(* IEC 61131-3 sources: plc-st-coding-agent/progress/evidence/f14_v10_full_20261113/jobs/codex_minimax-m27 (part 5) *)

(* ---- public-medium-04.candidate_04.st ---- *)
(* CONTRACT_RULES [] *)
FUNCTION_BLOCK FB_TemperatureControl
VAR_INPUT
    TemperatureSensorInput : REAL;
    SetTemperature         : REAL;
END_VAR
VAR_OUTPUT
    CurrentTemperature : REAL;
    SetTempDisplay      : REAL;
    HeaterStatus        : BOOL;
    OverheatProtection  : BOOL;
    HeaterOutput        : BOOL;
END_VAR
VAR
    tonCooldown         : TON;
    local_OverheatActive : BOOL := FALSE;
    local_SensorFault    : BOOL := FALSE;
    local_RuntimeAccum   : LTIME := LTIME#0s;
END_VAR

(* ENGINEERING_CONTRACT
  PUB003: Overheat protection triggers when heater runs continuously > 5s.
    - Activation: local_RuntimeAccum exceeds 5s on same scan it is detected.
    - Retention: OverheatActive stays TRUE until cooldown completes.
    - Reset/Deactivation: 3s cooldown via tonCooldown; heating condition
      must reassert AND cooldown must complete before heater can restart.
    - Same-scan priority: heater outputs set to FALSE when overheat activates;
      local_RuntimeAccum resets only when heating condition drops (not on
      overheat trigger), preserving correct accumulated-time logic.
    - Units/Boundaries: LTIME nanoseconds; strict > 5000ms threshold.
  PUB004: Heater turns on when temperature < setpoint (strict <).
  PUB007: Status outputs reflect current state every scan.
  PUB006: Sensor fault (input < 0 or > 100) turns heater off immediately.
*)

CurrentTemperature := TemperatureSensorInput;
SetTempDisplay     := SetTemperature;

local_SensorFault := (TemperatureSensorInput < 0.0) OR (TemperatureSensorInput > 100.0);

IF local_SensorFault OR local_OverheatActive THEN
    HeaterOutput := FALSE;
ELSE
    IF TemperatureSensorInput < SetTemperature THEN
        HeaterOutput := TRUE;
    ELSE
        HeaterOutput := FALSE;
    END_IF;
END_IF;

IF HeaterOutput THEN
    local_RuntimeAccum := local_RuntimeAccum + TO_LTIME(1);
END_IF;

IF NOT HeaterOutput THEN
    local_RuntimeAccum := LTIME#0s;
END_IF;

IF local_RuntimeAccum > T#5s THEN
    local_OverheatActive := TRUE;
    local_RuntimeAccum   := LTIME#0s;
END_IF;

IF local_OverheatActive THEN
    tonCooldown(IN := TRUE, PT := T#3s);
    IF tonCooldown.Q THEN
        local_OverheatActive := FALSE;
    END_IF;
ELSE
    tonCooldown(IN := FALSE, PT := T#3s);
END_IF;

HeaterStatus       := HeaterOutput;
OverheatProtection := local_OverheatActive;
END_FUNCTION_BLOCK

(* ---- public-medium-04.raw_candidate_01.st ---- *)
(*
ENGINEERING_CONTRACT:
PUB001: Read TemperatureSensorInput (REAL), display in CurrentTemperature
PUB002: HeaterOutput := TRUE when TemperatureSensorInput < SetTemperature
PUB003: Overheat triggers after >5s continuous HeaterOutput (strict > boundary)
PUB004: Overheat auto-sets HeaterOutput:=FALSE, 3s cooldown before OverheatProtection can clear
PUB005: Sensor fault (<0 OR >100) sets HeaterOutput:=FALSE regardless of temperature
PUB006: Status outputs (CurrentTemperature, SetTempDisplay, HeaterStatus, OverheatProtection) update every scan

Activation: All outputs update every scan (no edge-only behavior)
Retention: OverheatActive retains state across scans until cooldown completes
Reset/Deactivation: OverheatActive resets only after OverheatCooldownTimer.Q (3s elapsed)
Same-scan priority: HeaterOutput finalized BEFORE runtime timer enable is evaluated
Units: TIME/LTIME for timers (TON), REAL for temperatures, BOOL for control/status
*)
FUNCTION_BLOCK FB_TemperatureControl
VAR_INPUT
    TemperatureSensorInput : REAL;
    SetTemperature : REAL;
END_VAR

VAR_OUTPUT
    CurrentTemperature : REAL;
    SetTempDisplay : REAL;
    HeaterStatus : BOOL;
    OverheatProtection : BOOL;
    HeaterOutput : BOOL;
END_VAR

VAR
    HeaterRuntimeTimer : TON;
    OverheatCooldownTimer : TON;
    OverheatActive : BOOL := FALSE;
    SensorFault : BOOL := FALSE;
END_VAR

// Update display outputs
CurrentTemperature := TemperatureSensorInput;
SetTempDisplay := SetTemperature;

// Sensor fault detection: invalid range turns off heater
SensorFault := (TemperatureSensorInput < 0.0) OR (TemperatureSensorInput > 100.0);

// Temperature control logic
IF NOT SensorFault AND NOT OverheatActive THEN
    // Normal operation: heater ON when below setpoint
    IF TemperatureSensorInput < SetTemperature THEN
        HeaterOutput := TRUE;
    ELSE
        HeaterOutput := FALSE;
    END_IF;
ELSE
    // Sensor fault or overheat protection active - heater OFF
    HeaterOutput := FALSE;
END_IF;

// Update heater status display
HeaterStatus := HeaterOutput;

// Runtime timer: tracks continuous heater ON time (resets when heater OFF)
HeaterRuntimeTimer(IN := HeaterOutput, PT := T#5s);

// Overheat detection: >5s continuous heater operation
IF HeaterRuntimeTimer.Q AND NOT OverheatActive THEN
    OverheatActive := TRUE;
    OverheatCooldownTimer(IN := TRUE, PT := T#3s);
END_IF;

// Overheat cooldown: 3s wait before protection can be lifted
IF OverheatActive THEN
    OverheatCooldownTimer(IN := TRUE, PT := T#3s);
    IF OverheatCooldownTimer.Q THEN
        OverheatActive := FALSE;
    END_IF;
END_IF;

// Update overheat protection status
OverheatProtection := OverheatActive;
END_FUNCTION_BLOCK

(* ---- public-medium-04.raw_candidate_02.st ---- *)
(*
ENGINEERING_CONTRACT:
PUB001: TemperatureSensorInput (REAL) -> CurrentTemperature (REAL) every scan
PUB002: HeaterOutput := TRUE when TemperatureSensorInput < SetTemperature (no sensor fault)
PUB003: Overheat triggers when runtime > 5s (strict >), first satisfying tick = 5001ms
PUB004: Overheat sets HeaterOutput:=FALSE, 3s cooldown before OverheatProtection clears
PUB005: Sensor fault (<0 OR >100) sets HeaterOutput:=FALSE regardless of temperature
PUB006: All status outputs (CurrentTemperature, SetTempDisplay, HeaterStatus, OverheatProtection) update every scan
*)
FUNCTION_BLOCK FB_TemperatureControl
VAR_INPUT
    TemperatureSensorInput : REAL;
    SetTemperature         : REAL;
END_VAR

VAR_OUTPUT
    CurrentTemperature : REAL;
    SetTempDisplay      : REAL;
    HeaterStatus        : BOOL;
    OverheatProtection  : BOOL;
    HeaterOutput        : BOOL;
END_VAR

VAR
    HeaterRuntimeTimer   : TON;
    OverheatCooldownTimer: TON;
    OverheatActive       : BOOL := FALSE;
    SensorFault          : BOOL := FALSE;
    Runtimems            : LINT := 0;
END_VAR

SensorFault := (TemperatureSensorInput < 0.0) OR (TemperatureSensorInput > 100.0);

IF NOT SensorFault AND NOT OverheatActive THEN
    IF TemperatureSensorInput < SetTemperature THEN
        HeaterOutput := TRUE;
    ELSE
        HeaterOutput := FALSE;
    END_IF;
ELSE
    HeaterOutput := FALSE;
END_IF;

HeaterRuntimeTimer(IN := FALSE, PT := T#5s);

IF OverheatActive THEN
    IF Runtimems > 5000 THEN
        OverheatActive := TRUE;
    END_IF;
ELSIF HeaterOutput THEN
    Runtimems := Runtimems + TO_LINT(HeaterRuntimeTimer.ET) + 1;
    HeaterRuntimeTimer(IN := TRUE, PT := T#5s);
    IF Runtimems > 5000 THEN
        OverheatActive := TRUE;
        HeaterOutput := FALSE;
    END_IF;
ELSE
    Runtimems := 0;
END_IF;

IF OverheatActive THEN
    OverheatCooldownTimer(IN := TRUE, PT := T#3s);
    IF OverheatCooldownTimer.Q THEN
        OverheatActive := FALSE;
        Runtimems := 0;
    END_IF;
END_IF;

CurrentTemperature := TemperatureSensorInput;
SetTempDisplay := SetTemperature;
HeaterStatus := HeaterOutput;
OverheatProtection := OverheatActive;
END_FUNCTION_BLOCK

(* ---- public-medium-04.raw_candidate_03.st ---- *)
(* CONTRACT_RULES [] *)
FUNCTION_BLOCK FB_TemperatureControl
VAR_INPUT
    TemperatureSensorInput : REAL;
    SetTemperature : REAL;
END_VAR
VAR_OUTPUT
    CurrentTemperature : REAL;
    SetTempDisplay : REAL;
    HeaterStatus : BOOL;
    OverheatProtection : BOOL;
    HeaterOutput : BOOL;
END_VAR
VAR
    HeaterRuntimeTimer : TON;
    OverheatCooldownTimer : TON;
    OverheatActive : BOOL := FALSE;
    SensorFault : BOOL := FALSE;
END_VAR

CurrentTemperature := TemperatureSensorInput;
SetTempDisplay := SetTemperature;
SensorFault := (TemperatureSensorInput < 0.0) OR (TemperatureSensorInput > 100.0);

HeaterRuntimeTimer(IN := (TemperatureSensorInput < SetTemperature) AND NOT SensorFault AND NOT OverheatActive, PT := T#5s);

IF HeaterRuntimeTimer.Q AND NOT OverheatActive THEN
    OverheatActive := TRUE;
    OverheatCooldownTimer(IN := TRUE, PT := T#3s);
END_IF;

IF OverheatActive THEN
    OverheatCooldownTimer(IN := TRUE, PT := T#3s);
    IF OverheatCooldownTimer.Q THEN
        OverheatActive := FALSE;
    END_IF;
END_IF;

IF NOT SensorFault AND NOT OverheatActive THEN
    IF TemperatureSensorInput < SetTemperature THEN
        HeaterOutput := TRUE;
    ELSE
        HeaterOutput := FALSE;
    END_IF;
ELSE
    HeaterOutput := FALSE;
END_IF;

HeaterStatus := HeaterOutput;
OverheatProtection := OverheatActive;
END_FUNCTION_BLOCK

(* ---- public-medium-04.raw_candidate_04.st ---- *)
(* CONTRACT_RULES [] *)
FUNCTION_BLOCK FB_TemperatureControl
VAR_INPUT
    TemperatureSensorInput : REAL;
    SetTemperature         : REAL;
END_VAR
VAR_OUTPUT
    CurrentTemperature : REAL;
    SetTempDisplay      : REAL;
    HeaterStatus        : BOOL;
    OverheatProtection  : BOOL;
    HeaterOutput        : BOOL;
END_VAR
VAR
    tonCooldown         : TON;
    local_OverheatActive : BOOL := FALSE;
    local_SensorFault    : BOOL := FALSE;
    local_RuntimeAccum   : LTIME := LTIME#0s;
END_VAR

(* ENGINEERING_CONTRACT
  PUB003: Overheat protection triggers when heater runs continuously > 5s.
    - Activation: local_RuntimeAccum exceeds 5s on same scan it is detected.
    - Retention: OverheatActive stays TRUE until cooldown completes.
    - Reset/Deactivation: 3s cooldown via tonCooldown; heating condition
      must reassert AND cooldown must complete before heater can restart.
    - Same-scan priority: heater outputs set to FALSE when overheat activates;
      local_RuntimeAccum resets only when heating condition drops (not on
      overheat trigger), preserving correct accumulated-time logic.
    - Units/Boundaries: LTIME nanoseconds; strict > 5000ms threshold.
  PUB004: Heater turns on when temperature < setpoint (strict <).
  PUB007: Status outputs reflect current state every scan.
  PUB006: Sensor fault (input < 0 or > 100) turns heater off immediately.
*)

CurrentTemperature := TemperatureSensorInput;
SetTempDisplay     := SetTemperature;

local_SensorFault := (TemperatureSensorInput < 0.0) OR (TemperatureSensorInput > 100.0);

IF local_SensorFault OR local_OverheatActive THEN
    HeaterOutput := FALSE;
ELSE
    IF TemperatureSensorInput < SetTemperature THEN
        HeaterOutput := TRUE;
    ELSE
        HeaterOutput := FALSE;
    END_IF;
END_IF;

IF HeaterOutput THEN
    local_RuntimeAccum := local_RuntimeAccum + TO_LTIME(1);
END_IF;

IF NOT HeaterOutput THEN
    local_RuntimeAccum := LTIME#0s;
END_IF;

IF local_RuntimeAccum > T#5s THEN
    local_OverheatActive := TRUE;
    local_RuntimeAccum   := LTIME#0s;
END_IF;

IF local_OverheatActive THEN
    tonCooldown(IN := TRUE, PT := T#3s);
    IF tonCooldown.Q THEN
        local_OverheatActive := FALSE;
    END_IF;
ELSE
    tonCooldown(IN := FALSE, PT := T#3s);
END_IF;

HeaterStatus       := HeaterOutput;
OverheatProtection := local_OverheatActive;
END_FUNCTION_BLOCK

(* ---- public-medium-05.candidate_01.st ---- *)
(* ENGINEERING_CONTRACT *)
(*
  | Output/State Group       | Activation                                  | Retention                    | Reset/Deactivation            | Same-Scan Priority | Units/Boundaries |
  |--------------------------|---------------------------------------------|------------------------------|-------------------------------|--------------------|------------------|
  | MotorForward (Auto)      | State<>IDLE AND Mode=1                      | Hold until State=IDLE        | State=IDLE OR Mode=0          | Same-scan          | PUB001,PUB007    |
  | MotorReverse (Manual)    | ForwardButton=1 AND Mode=0 AND ReverseButton=0 | Hold until condition false | ForwardButton=0 OR Mode=1   | Same-scan          | PUB006,PUB002    |
  | CompletionLight          | State=DONE AND SensorC=1 AND Mode=1         | Hold while SensorC=1         | SensorC=0 OR Mode=0           | Same-scan          | PUB004,PUB008    |
  | State: IDLE→A            | SensorA=1 AND Mode=1 AND State=IDLE         | Until next transition        | SensorC=0 (product removed)   | Same-scan          | PUB003           |
  | State: A→B               | ButtonA=1 AND State=A                       | Until next transition        | SensorC=0                      | Same-scan          | PUB003           |
  | State: B→C               | SensorB=1 AND State=B                       | Until next transition        | SensorC=0                      | Same-scan          | PUB003           |
  | State: C→DONE            | ButtonC=1 AND State=C                       | Until SensorC=0              | SensorC=0                      | Same-scan          | PUB003           |
*)
(* CONTRACT_RULES [] *)
FUNCTION_BLOCK ProductionLineControl
VAR_INPUT
    Mode : BOOL;
    ForwardButton : BOOL;
    ReverseButton : BOOL;
    SensorA : BOOL;
    SensorB : BOOL;
    SensorC : BOOL;
    ButtonA : BOOL;
    ButtonB : BOOL;
    ButtonC : BOOL;
END_VAR
VAR_OUTPUT
    MotorForward : BOOL;
    MotorReverse : BOOL;
    CompletionLight : BOOL;
END_VAR
VAR
    State : INT;
    IDLE : INT := 0;
    StateA : INT := 1;
    StateB : INT := 2;
    StateC : INT := 3;
    StateD : INT := 4;
END_VAR
    IF Mode = FALSE THEN
        State := IDLE;
    ELSIF Mode = TRUE THEN
        IF State = IDLE AND SensorA THEN
            State := StateA;
        ELSIF State = StateA AND ButtonA THEN
            State := StateB;
        ELSIF State = StateB AND SensorB THEN
            State := StateC;
        ELSIF State = StateC AND ButtonC THEN
            State := StateD;
        END_IF;
    END_IF;
    MotorForward := ((State <> IDLE) AND Mode) OR (ForwardButton AND (NOT Mode) AND (NOT ReverseButton));
    MotorReverse := ReverseButton AND (NOT Mode) AND (NOT ForwardButton);
    CompletionLight := (State = StateD) AND SensorC AND Mode;
END_FUNCTION_BLOCK

(* ---- public-medium-05.candidate_02.st ---- *)
(* ENGINEERING_CONTRACT *)
(*
  | Output/State Group       | Activation                                  | Retention                    | Reset/Deactivation            | Same-Scan Priority | Units/Boundaries |
  |--------------------------|---------------------------------------------|------------------------------|-------------------------------|--------------------|------------------|
  | MotorForward (Auto)      | State=B OR State=D_transit                  | Hold via tmp_MotorRunning    | State=C/DONE OR Mode=0         | Same-scan          | PUB006           |
  | MotorReverse (Manual)    | ReverseButton AND Mode=0 AND !ForwardButton | Hold until condition false   | !ReverseButton OR Mode=1       | Same-scan          | PUB004,PUB002    |
  | CompletionLight          | State=DONE AND SensorC AND Mode             | Hold while SensorC           | SensorC=0 OR Mode=0            | Same-scan          | PUB008           |
  | State transitions        | Per clause PUB003                           | Until next trigger           | Mode=0 → IDLE                  | Same-scan          | PUB003           |
*)
(* CONTRACT_RULES [] *)
FUNCTION_BLOCK ProductionLineControl
VAR_INPUT
    Mode : BOOL;
    ForwardButton : BOOL;
    ReverseButton : BOOL;
    SensorA : BOOL;
    SensorB : BOOL;
    SensorC : BOOL;
    ButtonA : BOOL;
    ButtonB : BOOL;
    ButtonC : BOOL;
END_VAR
VAR_OUTPUT
    MotorForward : BOOL;
    MotorReverse : BOOL;
    CompletionLight : BOOL;
END_VAR
VAR
    State : INT;
    IDLE : INT := 0;
    StateA : INT := 1;
    StateB : INT := 2;
    StateC : INT := 3;
    StateD_transit : INT := 4;
    DONE : INT := 5;
    tmp_MotorRunning : BOOL;
END_VAR
    tmp_MotorRunning := (State = StateB) OR (State = StateD_transit);
    MotorForward := tmp_MotorRunning AND Mode;
    MotorReverse := ReverseButton AND (NOT Mode) AND (NOT ForwardButton);
    CompletionLight := (State = DONE) AND SensorC AND Mode;
    IF Mode = FALSE THEN
        State := IDLE;
    ELSIF Mode = TRUE THEN
        IF State = IDLE AND SensorA THEN
            State := StateA;
        ELSIF State = StateA AND ButtonA THEN
            State := StateB;
            tmp_MotorRunning := TRUE;
        ELSIF State = StateB AND SensorB THEN
            State := StateC;
        ELSIF State = StateC AND ButtonC THEN
            State := StateD_transit;
            tmp_MotorRunning := TRUE;
        ELSIF State = StateD_transit AND SensorC THEN
            State := DONE;
        ELSIF State = DONE AND NOT SensorC THEN
            State := IDLE;
        END_IF;
    END_IF;
END_FUNCTION_BLOCK

(* ---- public-medium-05.candidate_03.st ---- *)
(* ENGINEERING_CONTRACT *)
(*
  | Output/State Group       | Activation                                  | Retention                    | Reset/Deactivation            | Same-Scan Priority | Units/Boundaries |
  |--------------------------|---------------------------------------------|------------------------------|-------------------------------|--------------------|------------------|
  | MotorForward (Auto)      | State=StateA OR State=StateB AND Mode=1      | Hold until State=C or IDLE   | State=C/D OR Mode=0          | Same-scan          | PUB001,PUB007    |
  | MotorReverse (Manual)    | ForwardButton=1 AND Mode=0 AND ReverseButton=0 | Hold until condition false | ForwardButton=0 OR Mode=1   | Same-scan          | PUB006,PUB002    |
  | CompletionLight          | State=StateD AND SensorC=1 AND Mode=1        | Hold while SensorC=1         | SensorC=0 OR Mode=0           | Same-scan          | PUB004,PUB008    |
  | State: IDLE→A            | SensorA=1 AND Mode=1 AND State=IDLE          | Until next transition        | SensorC=0 (product removed)   | Same-scan          | PUB003           |
  | State: A→B               | ButtonA=1 AND State=StateA                   | Until next transition        | SensorC=0                     | Same-scan          | PUB003           |
  | State: B→C               | SensorB=1 AND State=StateB                   | Until next transition        | SensorC=0                     | Same-scan          | PUB003           |
  | State: C→DONE            | ButtonC=1 AND State=StateC                   | Until SensorC=0              | SensorC=0                     | Same-scan          | PUB003           |
*)
(* CONTRACT_RULES [] *)
FUNCTION_BLOCK ProductionLineControl
VAR_INPUT
    Mode : BOOL;
    ForwardButton : BOOL;
    ReverseButton : BOOL;
    SensorA : BOOL;
    SensorB : BOOL;
    SensorC : BOOL;
    ButtonA : BOOL;
    ButtonB : BOOL;
    ButtonC : BOOL;
END_VAR
VAR_OUTPUT
    MotorForward : BOOL;
    MotorReverse : BOOL;
    CompletionLight : BOOL;
END_VAR
VAR
    State : INT;
    IDLE : INT := 0;
    StateA : INT := 1;
    StateB : INT := 2;
    StateC : INT := 3;
    StateD : INT := 4;
END_VAR
    IF Mode = FALSE THEN
        State := IDLE;
    ELSIF Mode = TRUE THEN
        IF State = IDLE AND SensorA THEN
            State := StateA;
        ELSIF State = StateA AND ButtonA THEN
            State := StateB;
        ELSIF State = StateB AND SensorB THEN
            State := StateC;
        ELSIF State = StateC AND ButtonC THEN
            State := StateD;
        END_IF;
    END_IF;
    MotorForward := ((State = StateA) OR (State = StateB)) AND Mode OR (ForwardButton AND (NOT Mode) AND (NOT ReverseButton));
    MotorReverse := ReverseButton AND (NOT Mode) AND (NOT ForwardButton);
    CompletionLight := (State = StateD) AND SensorC AND Mode;
END_FUNCTION_BLOCK

(* ---- public-medium-05.candidate_04.st ---- *)
(* ENGINEERING_CONTRACT *)
(*
  | Output/State Group       | Activation                                  | Retention                    | Reset/Deactivation            | Same-Scan Priority | Units/Boundaries |
  |--------------------------|---------------------------------------------|------------------------------|-------------------------------|--------------------|------------------|
  | MotorForward (Auto)      | State=A/B/D AND Mode=1                      | Hold until State=IDLE        | Mode=0 OR State=IDLE          | Same-scan          | PUB001,PUB007    |
  | MotorForward (Manual)    | ForwardButton=1 AND Mode=0 AND ReverseButton=0 | Hold until condition false | ForwardButton=0 OR Mode=1   | Same-scan          | PUB006,PUB002    |
  | CompletionLight          | State=StateD AND SensorC=1 AND Mode=1        | Hold while SensorC=1         | SensorC=0 OR Mode=0           | Same-scan          | PUB004,PUB008    |
  | State: IDLE→A            | SensorA=1 AND Mode=1 AND State=IDLE          | Until next transition        | SensorC=0 (product removed)   | Same-scan          | PUB003           |
  | State: A→B               | ButtonA=1 AND State=StateA                   | Until next transition        | SensorC=0                     | Same-scan          | PUB003           |
  | State: B→C               | SensorB=1 AND State=StateB                   | Until next transition        | SensorC=0                     | Same-scan          | PUB003           |
  | State: C→DONE            | ButtonC=1 AND State=StateC                   | Until SensorC=0              | SensorC=0                     | Same-scan          | PUB003           |
*)
(* CONTRACT_RULES [] *)
FUNCTION_BLOCK ProductionLineControl
VAR_INPUT
    Mode : BOOL;
    ForwardButton : BOOL;
    ReverseButton : BOOL;
    SensorA : BOOL;
    SensorB : BOOL;
    SensorC : BOOL;
    ButtonA : BOOL;
    ButtonB : BOOL;
    ButtonC : BOOL;
END_VAR
VAR_OUTPUT
    MotorForward : BOOL;
    MotorReverse : BOOL;
    CompletionLight : BOOL;
END_VAR
VAR
    State : INT;
    IDLE : INT := 0;
    StateA : INT := 1;
    StateB : INT := 2;
    StateC : INT := 3;
    StateD : INT := 4;
END_VAR
    IF Mode = FALSE THEN
        State := IDLE;
    ELSIF Mode = TRUE THEN
        IF State = IDLE AND SensorA THEN
            State := StateA;
        ELSIF State = StateA AND ButtonA THEN
            State := StateB;
        ELSIF State = StateB AND SensorB THEN
            State := StateC;
        ELSIF State = StateC AND ButtonC THEN
            State := StateD;
        END_IF;
    END_IF;
    MotorForward := ((State = StateA) OR (State = StateB) OR (State = StateD)) AND Mode OR (ForwardButton AND (NOT Mode) AND (NOT ReverseButton));
    MotorReverse := ReverseButton AND (NOT Mode) AND (NOT ForwardButton);
    CompletionLight := (State = StateD) AND SensorC AND Mode;
END_FUNCTION_BLOCK

(* ---- public-medium-05.raw_candidate_01.st ---- *)
(* ENGINEERING_CONTRACT *)
(*
  | Output/State Group       | Activation                                  | Retention                    | Reset/Deactivation            | Same-Scan Priority | Units/Boundaries |
  |--------------------------|---------------------------------------------|------------------------------|-------------------------------|--------------------|------------------|
  | MotorForward (Auto)      | State<>IDLE AND Mode=1                      | Hold until State=IDLE        | State=IDLE OR Mode=0          | Same-scan          | PUB001,PUB007    |
  | MotorReverse (Manual)    | ForwardButton=1 AND Mode=0 AND ReverseButton=0 | Hold until condition false | ForwardButton=0 OR Mode=1   | Same-scan          | PUB006,PUB002    |
  | CompletionLight          | State=DONE AND SensorC=1 AND Mode=1         | Hold while SensorC=1         | SensorC=0 OR Mode=0           | Same-scan          | PUB004,PUB008    |
  | State: IDLE→A            | SensorA=1 AND Mode=1 AND State=IDLE         | Until next transition        | SensorC=0 (product removed)   | Same-scan          | PUB003           |
  | State: A→B               | ButtonA=1 AND State=A                       | Until next transition        | SensorC=0                      | Same-scan          | PUB003           |
  | State: B→C               | SensorB=1 AND State=B                       | Until next transition        | SensorC=0                      | Same-scan          | PUB003           |
  | State: C→DONE            | ButtonC=1 AND State=C                       | Until SensorC=0              | SensorC=0                      | Same-scan          | PUB003           |
*)
(* CONTRACT_RULES [] *)
FUNCTION_BLOCK ProductionLineControl
VAR_INPUT
    Mode : BOOL;
    ForwardButton : BOOL;
    ReverseButton : BOOL;
    SensorA : BOOL;
    SensorB : BOOL;
    SensorC : BOOL;
    ButtonA : BOOL;
    ButtonB : BOOL;
    ButtonC : BOOL;
END_VAR
VAR_OUTPUT
    MotorForward : BOOL;
    MotorReverse : BOOL;
    CompletionLight : BOOL;
END_VAR
VAR
    State : INT;
    IDLE : INT := 0;
    StateA : INT := 1;
    StateB : INT := 2;
    StateC : INT := 3;
    StateD : INT := 4;
END_VAR
    IF Mode = FALSE THEN
        State := IDLE;
    ELSIF Mode = TRUE THEN
        IF State = IDLE AND SensorA THEN
            State := StateA;
        ELSIF State = StateA AND ButtonA THEN
            State := StateB;
        ELSIF State = StateB AND SensorB THEN
            State := StateC;
        ELSIF State = StateC AND ButtonC THEN
            State := StateD;
        END_IF;
    END_IF;
    MotorForward := ((State <> IDLE) AND Mode) OR (ForwardButton AND (NOT Mode) AND (NOT ReverseButton));
    MotorReverse := ReverseButton AND (NOT Mode) AND (NOT ForwardButton);
    CompletionLight := (State = StateD) AND SensorC AND Mode;
END_FUNCTION_BLOCK

(* ---- public-medium-05.raw_candidate_02.st ---- *)
(* ENGINEERING_CONTRACT *)
(*
  | Output/State Group       | Activation                                  | Retention                    | Reset/Deactivation            | Same-Scan Priority | Units/Boundaries |
  |--------------------------|---------------------------------------------|------------------------------|-------------------------------|--------------------|------------------|
  | MotorForward (Auto)      | State=B OR State=D_transit                  | Hold via tmp_MotorRunning    | State=C/DONE OR Mode=0         | Same-scan          | PUB006           |
  | MotorReverse (Manual)    | ReverseButton AND Mode=0 AND !ForwardButton | Hold until condition false   | !ReverseButton OR Mode=1       | Same-scan          | PUB004,PUB002    |
  | CompletionLight          | State=DONE AND SensorC AND Mode             | Hold while SensorC           | SensorC=0 OR Mode=0            | Same-scan          | PUB008           |
  | State transitions        | Per clause PUB003                           | Until next trigger           | Mode=0 → IDLE                  | Same-scan          | PUB003           |
*)
(* CONTRACT_RULES [] *)
FUNCTION_BLOCK ProductionLineControl
VAR_INPUT
    Mode : BOOL;
    ForwardButton : BOOL;
    ReverseButton : BOOL;
    SensorA : BOOL;
    SensorB : BOOL;
    SensorC : BOOL;
    ButtonA : BOOL;
    ButtonB : BOOL;
    ButtonC : BOOL;
END_VAR
VAR_OUTPUT
    MotorForward : BOOL;
    MotorReverse : BOOL;
    CompletionLight : BOOL;
END_VAR
VAR
    State : INT;
    IDLE : INT := 0;
    StateA : INT := 1;
    StateB : INT := 2;
    StateC : INT := 3;
    StateD_transit : INT := 4;
    DONE : INT := 5;
    tmp_MotorRunning : BOOL;
END_VAR
    tmp_MotorRunning := (State = StateB) OR (State = StateD_transit);
    MotorForward := tmp_MotorRunning AND Mode;
    MotorReverse := ReverseButton AND (NOT Mode) AND (NOT ForwardButton);
    CompletionLight := (State = DONE) AND SensorC AND Mode;
    IF Mode = FALSE THEN
        State := IDLE;
    ELSIF Mode = TRUE THEN
        IF State = IDLE AND SensorA THEN
            State := StateA;
        ELSIF State = StateA AND ButtonA THEN
            State := StateB;
            tmp_MotorRunning := TRUE;
        ELSIF State = StateB AND SensorB THEN
            State := StateC;
        ELSIF State = StateC AND ButtonC THEN
            State := StateD_transit;
            tmp_MotorRunning := TRUE;
        ELSIF State = StateD_transit AND SensorC THEN
            State := DONE;
        ELSIF State = DONE AND NOT SensorC THEN
            State := IDLE;
        END_IF;
    END_IF;
END_FUNCTION_BLOCK

(* ---- public-medium-05.raw_candidate_03.st ---- *)
(* ENGINEERING_CONTRACT *)
(*
  | Output/State Group       | Activation                                  | Retention                    | Reset/Deactivation            | Same-Scan Priority | Units/Boundaries |
  |--------------------------|---------------------------------------------|------------------------------|-------------------------------|--------------------|------------------|
  | MotorForward (Auto)      | State=StateA OR State=StateB AND Mode=1      | Hold until State=C or IDLE   | State=C/D OR Mode=0          | Same-scan          | PUB001,PUB007    |
  | MotorReverse (Manual)    | ForwardButton=1 AND Mode=0 AND ReverseButton=0 | Hold until condition false | ForwardButton=0 OR Mode=1   | Same-scan          | PUB006,PUB002    |
  | CompletionLight          | State=StateD AND SensorC=1 AND Mode=1        | Hold while SensorC=1         | SensorC=0 OR Mode=0           | Same-scan          | PUB004,PUB008    |
  | State: IDLE→A            | SensorA=1 AND Mode=1 AND State=IDLE          | Until next transition        | SensorC=0 (product removed)   | Same-scan          | PUB003           |
  | State: A→B               | ButtonA=1 AND State=StateA                   | Until next transition        | SensorC=0                     | Same-scan          | PUB003           |
  | State: B→C               | SensorB=1 AND State=StateB                   | Until next transition        | SensorC=0                     | Same-scan          | PUB003           |
  | State: C→DONE            | ButtonC=1 AND State=StateC                   | Until SensorC=0              | SensorC=0                     | Same-scan          | PUB003           |
*)
(* CONTRACT_RULES [] *)
FUNCTION_BLOCK ProductionLineControl
VAR_INPUT
    Mode : BOOL;
    ForwardButton : BOOL;
    ReverseButton : BOOL;
    SensorA : BOOL;
    SensorB : BOOL;
    SensorC : BOOL;
    ButtonA : BOOL;
    ButtonB : BOOL;
    ButtonC : BOOL;
END_VAR
VAR_OUTPUT
    MotorForward : BOOL;
    MotorReverse : BOOL;
    CompletionLight : BOOL;
END_VAR
VAR
    State : INT;
    IDLE : INT := 0;
    StateA : INT := 1;
    StateB : INT := 2;
    StateC : INT := 3;
    StateD : INT := 4;
END_VAR
    IF Mode = FALSE THEN
        State := IDLE;
    ELSIF Mode = TRUE THEN
        IF State = IDLE AND SensorA THEN
            State := StateA;
        ELSIF State = StateA AND ButtonA THEN
            State := StateB;
        ELSIF State = StateB AND SensorB THEN
            State := StateC;
        ELSIF State = StateC AND ButtonC THEN
            State := StateD;
        END_IF;
    END_IF;
    MotorForward := ((State = StateA) OR (State = StateB)) AND Mode OR (ForwardButton AND (NOT Mode) AND (NOT ReverseButton));
    MotorReverse := ReverseButton AND (NOT Mode) AND (NOT ForwardButton);
    CompletionLight := (State = StateD) AND SensorC AND Mode;
END_FUNCTION_BLOCK

(* ---- public-medium-05.raw_candidate_04.st ---- *)
(* ENGINEERING_CONTRACT *)
(*
  | Output/State Group       | Activation                                  | Retention                    | Reset/Deactivation            | Same-Scan Priority | Units/Boundaries |
  |--------------------------|---------------------------------------------|------------------------------|-------------------------------|--------------------|------------------|
  | MotorForward (Auto)      | State=A/B/D AND Mode=1                      | Hold until State=IDLE        | Mode=0 OR State=IDLE          | Same-scan          | PUB001,PUB007    |
  | MotorForward (Manual)    | ForwardButton=1 AND Mode=0 AND ReverseButton=0 | Hold until condition false | ForwardButton=0 OR Mode=1   | Same-scan          | PUB006,PUB002    |
  | CompletionLight          | State=StateD AND SensorC=1 AND Mode=1        | Hold while SensorC=1         | SensorC=0 OR Mode=0           | Same-scan          | PUB004,PUB008    |
  | State: IDLE→A            | SensorA=1 AND Mode=1 AND State=IDLE          | Until next transition        | SensorC=0 (product removed)   | Same-scan          | PUB003           |
  | State: A→B               | ButtonA=1 AND State=StateA                   | Until next transition        | SensorC=0                     | Same-scan          | PUB003           |
  | State: B→C               | SensorB=1 AND State=StateB                   | Until next transition        | SensorC=0                     | Same-scan          | PUB003           |
  | State: C→DONE            | ButtonC=1 AND State=StateC                   | Until SensorC=0              | SensorC=0                     | Same-scan          | PUB003           |
*)
(* CONTRACT_RULES [] *)
FUNCTION_BLOCK ProductionLineControl
VAR_INPUT
    Mode : BOOL;
    ForwardButton : BOOL;
    ReverseButton : BOOL;
    SensorA : BOOL;
    SensorB : BOOL;
    SensorC : BOOL;
    ButtonA : BOOL;
    ButtonB : BOOL;
    ButtonC : BOOL;
END_VAR
VAR_OUTPUT
    MotorForward : BOOL;
    MotorReverse : BOOL;
    CompletionLight : BOOL;
END_VAR
VAR
    State : INT;
    IDLE : INT := 0;
    StateA : INT := 1;
    StateB : INT := 2;
    StateC : INT := 3;
    StateD : INT := 4;
END_VAR
    IF Mode = FALSE THEN
        State := IDLE;
    ELSIF Mode = TRUE THEN
        IF State = IDLE AND SensorA THEN
            State := StateA;
        ELSIF State = StateA AND ButtonA THEN
            State := StateB;
        ELSIF State = StateB AND SensorB THEN
            State := StateC;
        ELSIF State = StateC AND ButtonC THEN
            State := StateD;
        END_IF;
    END_IF;
    MotorForward := ((State = StateA) OR (State = StateB) OR (State = StateD)) AND Mode OR (ForwardButton AND (NOT Mode) AND (NOT ReverseButton));
    MotorReverse := ReverseButton AND (NOT Mode) AND (NOT ForwardButton);
    CompletionLight := (State = StateD) AND SensorC AND Mode;
END_FUNCTION_BLOCK

(* ---- public-medium-06.candidate_01.st ---- *)
FUNCTION_BLOCK SlabThicknessMonitor
VAR_INPUT
    THICKNESS_FAULT        : BOOL;
    THICKNESS_SIGNAL_VALID : BOOL;
    CUTTING_RUN            : BOOL;
    FaultTimestamp         : DINT;
    CycleTime              : TIME;
END_VAR

VAR_OUTPUT
    THICKNESS_ALARM          : BOOL;
    Slab_Fault_Counter       : UINT;
    Slab_Runtime_Accumulator : LTIME;
    Slab_Fault_History       : ARRAY[0..4] OF DINT;
END_VAR

VAR
    faultRising      : R_TRIG;
    validFalling     : R_TRIG;
    prevFault        : BOOL;
    prevValid        : BOOL;
    holdTimer        : TON;
    tmpI             : UINT;
END_VAR

(* ENGINEERING_CONTRACT
 * ┌─────────────────────────────────────────────────────────────────────────────────────────────┐
 * │ OUTPUT STATE TABLE                                                                           │
 * ├─────────────────┬───────────────────────────────────────────────────────────────────────────┤
 * │ THICKNESS_ALARM │ Activation:   rising edge of THICKNESS_FAULT while VALID=TRUE (PUB001)    │
 * │                 │ Retention:    held >= 500 ms via TON; remains TRUE while FAULT persists   │
 * │                 │ Reset:        VALID=FALSE or power-up clears alarm and holding state (PUB004)│
 * │                 │ Same-scan:    if VALID drops mid-scan, alarm OFF regardless of FAULT state│
 * ├─────────────────┼───────────────────────────────────────────────────────────────────────────┤
 * │ Slab_Fault_     │ Activation:   FALSE-to-TRUE of FAULT while VALID=TRUE (PUB002)             │
 * │ Counter         │ Retention:    monotonically increasing; never auto-decremented             │
 * │                 │ Reset:        power-up only (PUB005); external callers cannot modify       │
 * │                 │ Boundary:     UINT range; overflow wraps per IEC 61131-3                  │
 * ├─────────────────┼───────────────────────────────────────────────────────────────────────────┤
 * │ Slab_Runtime_   │ Activation:   CUTTING_RUN AND VALID AND NOT FAULT each scan (PUB003)       │
 * │ Accumulator     │ Retention:    preserved when conditions not met; never auto-cleared       │
 * │                 │ Reset:        power-up only (PUB005); uses LTIME nanoseconds internally   │
 * │                 │ Units:        CycleTime (TIME/ms) converted to LTIME (ns) before add      │
 * ├─────────────────┼───────────────────────────────────────────────────────────────────────────┤
 * │ Slab_Fault_     │ Activation:   new entry at index 0 on valid fault transition (PUB002)     │
 * │ History[0..4]   │ Shift:        older entries shift toward higher indices (PUB002)           │
 * │                 │ Retention:    five most recent; older beyond index 4 are discarded        │
 * │                 │ Reset:        power-up zeros all five entries (PUB005); read-only to callers│
 * └─────────────────┴───────────────────────────────────────────────────────────────────────────┘
 *
 * ┌─────────────────────────────────────────────────────────────────────────────────────────────┐
 * │ INPUT BEHAVIOR                                                                               │
 * ├───────────────────────────────┬─────────────────────────────────────────────────────────────┤
 * │ THICKNESS_SIGNAL_VALID=FALSE  │ alarm OFF, timer reset, no fault record, no runtime accum   │
 * │ THICKNESS_SIGNAL_VALID=TRUE   │ normal monitoring; alarm follows FAULT, counter/hist update │
 * │ CUTTING_RUN=FALSE             │ no runtime accumulation (fault monitoring still active)     │
 * │ CycleTime positive assumption │ caller guarantees > T#0s per task spec                     │
 * └───────────────────────────────┴─────────────────────────────────────────────────────────────┘
 *
 * ┌─────────────────────────────────────────────────────────────────────────────────────────────┐
 * │ TIMING BOUNDARY (PUB001, PUB003)                                                            │
 * │ - 500 ms hold: TON.Q = elapsed >= PT; first satisfying tick = ceil(500ms/1ms) = 500 ticks   │
 * │ - No implicit one-scan delay; timer enable and Q check occur in same invocation            │
 * └─────────────────────────────────────────────────────────────────────────────────────────────┘
 *
 * CONTRACT_RULES [{"kind": "hold_until_reset", "output": "THICKNESS_ALARM", "set_input": "THICKNESS_FAULT", "reset_input": null}]
 *)

(* Power-up initialization: handled by VAR initial values *)

(* Detect rising edge of fault while signal is valid *)
faultRising(CLK := THICKNESS_FAULT AND THICKNESS_SIGNAL_VALID AND NOT prevFault);

(* Detect falling edge of VALID to clear alarm and timer *)
validFalling(CLK := prevValid AND NOT THICKNESS_SIGNAL_VALID);

(* Handle signal invalidation: clear alarm and timer holding state *)
IF validFalling.Q THEN
    THICKNESS_ALARM := FALSE;
    holdTimer(IN := FALSE, PT := T#500ms);
END_IF;

(* When VALID is FALSE, ensure alarm and timer are cleared *)
IF NOT THICKNESS_SIGNAL_VALID THEN
    THICKNESS_ALARM := FALSE;
    holdTimer(IN := FALSE, PT := T#500ms);
END_IF;

(* Process fault: activate alarm and record history *)
IF faultRising.Q THEN
    (* Increment fault counter *)
    Slab_Fault_Counter := Slab_Fault_Counter + 1;

    (* Shift history: move entries toward higher indices *)
    FOR tmpI := 4 TO 1 BY -1 DO
        Slab_Fault_History[tmpI] := Slab_Fault_History[tmpI - 1];
    END_FOR;

    (* Store new fault timestamp at index 0 *)
    Slab_Fault_History[0] := FaultTimestamp;

    (* Activate alarm and start hold timer *)
    THICKNESS_ALARM := TRUE;
    holdTimer(IN := TRUE, PT := T#500ms);
END_IF;

(* Maintain alarm while fault persists (after initial 500ms hold) *)
IF holdTimer.Q THEN
    THICKNESS_ALARM := THICKNESS_FAULT AND THICKNESS_SIGNAL_VALID;
    holdTimer(IN := THICKNESS_ALARM, PT := T#500ms);
END_IF;

(* Accumulate runtime while cutting normally *)
IF CUTTING_RUN AND THICKNESS_SIGNAL_VALID AND NOT THICKNESS_FAULT THEN
    Slab_Runtime_Accumulator := Slab_Runtime_Accumulator + TO_LTIME(CycleTime);
END_IF;

(* Update previous state for edge detection on next scan *)
prevFault := THICKNESS_FAULT;
prevValid := THICKNESS_SIGNAL_VALID;

END_FUNCTION_BLOCK

(* ---- public-medium-06.candidate_02.st ---- *)
FUNCTION_BLOCK SlabThicknessMonitor
VAR_INPUT
    THICKNESS_FAULT        : BOOL;
    THICKNESS_SIGNAL_VALID : BOOL;
    CUTTING_RUN            : BOOL;
    FaultTimestamp         : DINT;
    CycleTime              : TIME;
END_VAR

VAR_OUTPUT
    THICKNESS_ALARM          : BOOL;
    Slab_Fault_Counter       : UINT;
    Slab_Runtime_Accumulator : LTIME;
    Slab_Fault_History       : ARRAY[0..4] OF DINT;
END_VAR

VAR
    faultRising : R_TRIG;
    prevFault   : BOOL;
    prevValid   : BOOL;
    holdTimer   : TON;
    tmpI        : UINT;
END_VAR

(* ENGINEERING_CONTRACT
 * ┌─────────────────────────────────────────────────────────────────────────────────────────────┐
 * │ OUTPUT STATE TABLE                                                                           │
 * ├─────────────────┬───────────────────────────────────────────────────────────────────────────┤
 * │ THICKNESS_ALARM │ Activation:   immediate on rising edge of FAULT while VALID=TRUE (PUB001) │
 * │                 │ Retention:    hold >= 500ms via TON after FAULT drops; persists if FAULT │
 * │                 │               remains TRUE                                                │
 * │                 │ Reset:        VALID=FALSE clears alarm and timer holding state (PUB004)   │
 * │                 │ Same-scan:    alarm OFF immediately when VALID drops                      │
 * ├─────────────────┼───────────────────────────────────────────────────────────────────────────┤
 * │ Slab_Fault_     │ Activation:   FALSE-to-TRUE of FAULT while VALID=TRUE (PUB002)            │
 * │ Counter         │ Retention:    monotonically increasing; never auto-decremented            │
 * │                 │ Reset:        power-up only (PUB005)                                      │
 * │                 │ Boundary:     UINT range                                                  │
 * ├─────────────────┼───────────────────────────────────────────────────────────────────────────┤
 * │ Slab_Runtime_   │ Activation:   CUTTING_RUN AND VALID AND NOT FAULT AND NOT faultRising     │
 * │ Accumulator     │               (excludes scan where fault just transitioned TRUE) (PUB003) │
 * │                 │ Retention:    preserved when conditions not met                           │
 * │                 │ Reset:        power-up only (PUB005)                                      │
 * │                 │ Units:        CycleTime converted to LTIME ns before add                  │
 * ├─────────────────┼───────────────────────────────────────────────────────────────────────────┤
 * │ Slab_Fault_     │ Activation:   new entry at index 0 on valid fault transition (PUB002)     │
 * │ History[0..4]   │ Shift:        older entries shift toward higher indices (PUB002)          │
 * │                 │ Retention:    five most recent; older beyond index 4 discarded            │
 * │                 │ Reset:        power-up zeros all five entries (PUB005)                    │
 * └─────────────────┴───────────────────────────────────────────────────────────────────────────┘
 *
 * ┌─────────────────────────────────────────────────────────────────────────────────────────────┐
 * │ TIMING BOUNDARY (PUB001)                                                                    │
 * │ - 500ms hold: TON.Q = elapsed >= PT; first satisfying tick = 500 ticks at 1ms quantum      │
 * │ - Alarm reactivates immediately via R_TRIG on same-scan FAULT transitions                  │
 * │ - Timer resets when alarm deactivates to prevent stale elapsed time                        │
 * └─────────────────────────────────────────────────────────────────────────────────────────────┘
 *
 * CONTRACT_RULES [{"kind": "hold_until_reset", "output": "THICKNESS_ALARM", "set_input": "THICKNESS_FAULT", "reset_input": null}]
 *)

(* Power-up initialization: VAR initial values handle zeroing *)

(* Detect rising edge of fault while signal is valid *)
faultRising(CLK := THICKNESS_FAULT AND THICKNESS_SIGNAL_VALID AND NOT prevFault);

(* Clear alarm and timer when signal becomes invalid *)
IF NOT THICKNESS_SIGNAL_VALID THEN
    THICKNESS_ALARM := FALSE;
    holdTimer(IN := FALSE, PT := T#500ms);
END_IF;

(* Activate alarm immediately on valid fault rising edge *)
IF faultRising.Q THEN
    THICKNESS_ALARM := TRUE;
    holdTimer(IN := TRUE, PT := T#500ms);
END_IF;

(* Maintain alarm while fault persists after initial hold *)
IF holdTimer.Q THEN
    THICKNESS_ALARM := THICKNESS_FAULT AND THICKNESS_SIGNAL_VALID;
    holdTimer(IN := THICKNESS_ALARM, PT := T#500ms);
END_IF;

(* Record fault: increment counter and shift history *)
IF faultRising.Q THEN
    Slab_Fault_Counter := Slab_Fault_Counter + 1;
    FOR tmpI := 4 TO 1 BY -1 DO
        Slab_Fault_History[tmpI] := Slab_Fault_History[tmpI - 1];
    END_FOR;
    Slab_Fault_History[0] := FaultTimestamp;
END_IF;

(* Accumulate runtime only while cutting normally (excludes fault-transition scan) *)
IF CUTTING_RUN AND THICKNESS_SIGNAL_VALID AND NOT THICKNESS_FAULT AND NOT faultRising.Q THEN
    Slab_Runtime_Accumulator := Slab_Runtime_Accumulator + TO_LTIME(CycleTime);
END_IF;

(* Update previous state for edge detection *)
prevFault := THICKNESS_FAULT;
prevValid := THICKNESS_SIGNAL_VALID;

END_FUNCTION_BLOCK

(* ---- public-medium-06.candidate_03.st ---- *)
FUNCTION_BLOCK SlabThicknessMonitor
VAR_INPUT
    THICKNESS_FAULT        : BOOL;
    THICKNESS_SIGNAL_VALID : BOOL;
    CUTTING_RUN            : BOOL;
    FaultTimestamp         : DINT;
    CycleTime              : TIME;
END_VAR

VAR_OUTPUT
    THICKNESS_ALARM          : BOOL;
    Slab_Fault_Counter       : UINT;
    Slab_Runtime_Accumulator : LTIME;
    Slab_Fault_History       : ARRAY[0..4] OF DINT;
END_VAR

VAR
    faultRising  : R_TRIG;
    validFalling : F_TRIG;
    prevFault    : BOOL;
    prevValid    : BOOL;
    holdTimer    : TON;
    latch        : BOOL;
    inHoldPhase  : BOOL;
    tmpI         : UINT;
END_VAR

(* ENGINEERING_CONTRACT
 * ┌─────────────────────────────────────────────────────────────────────────────────────────────┐
 * │ OUTPUT STATE TABLE                                                                           │
 * ├─────────────────┬───────────────────────────────────────────────────────────────────────────┤
 * │ THICKNESS_ALARM │ Activation:   immediate on rising edge of FAULT while VALID=TRUE (PUB001) │
 * │                 │ Retention:    held >= 500ms via TON; remains TRUE while FAULT persists   │
 * │                 │ Reset:        VALID=FALSE clears latch and timer (PUB004)                 │
 * │                 │ Same-scan:    latch set and timer started in same invocation as rising edge│
 * ├─────────────────┼───────────────────────────────────────────────────────────────────────────┤
 * │ Slab_Fault_     │ Activation:   FALSE-to-TRUE of FAULT while VALID=TRUE (PUB002)            │
 * │ Counter         │ Retention:    monotonically increasing; never auto-decremented            │
 * │                 │ Reset:        power-up only (PUB005)                                     │
 * │                 │ Boundary:     UINT range; overflow wraps per IEC 61131-3                 │
 * ├─────────────────┼───────────────────────────────────────────────────────────────────────────┤
 * │ Slab_Runtime_   │ Activation:   CUTTING_RUN AND VALID AND NOT FAULT each scan (PUB003)      │
 * │ Accumulator     │ Retention:    preserved when conditions not met; never auto-cleared      │
 * │                 │ Reset:        power-up only (PUB005)                                     │
 * │                 │ Units:        CycleTime (TIME) converted to LTIME (ns) before add        │
 * ├─────────────────┼───────────────────────────────────────────────────────────────────────────┤
 * │ Slab_Fault_     │ Activation:   new entry at index 0 on valid fault transition (PUB002)    │
 * │ History[0..4]   │ Shift:        older entries shift toward higher indices (PUB002)          │
 * │                 │ Retention:    five most recent; older beyond index 4 are discarded       │
 * │                 │ Reset:        power-up zeros all five entries (PUB005)                   │
 * └─────────────────┴───────────────────────────────────────────────────────────────────────────┘
 *
 * ┌─────────────────────────────────────────────────────────────────────────────────────────────┐
 * │ TIMING BOUNDARY (PUB001)                                                                    │
 * │ - 500 ms hold: TON.Q = elapsed >= PT; first satisfying tick = ceil(500ms/1ms) = 500 ticks  │
 * │ - Timer reset before restart ensures deterministic restart behavior                        │
 * └─────────────────────────────────────────────────────────────────────────────────────────────┘
 *
 * CONTRACT_RULES [{"kind": "hold_until_reset", "output": "THICKNESS_ALARM", "set_input": "THICKNESS_FAULT", "reset_input": null}]
 *)

(* Detect rising edge of fault while signal is valid *)
faultRising(CLK := THICKNESS_FAULT AND THICKNESS_SIGNAL_VALID AND NOT prevFault);

(* Detect falling edge of VALID to clear state *)
validFalling(CLK := prevValid AND NOT THICKNESS_SIGNAL_VALID);

(* Handle signal invalidation: clear latch, alarm, and timer *)
IF validFalling.Q THEN
    latch := FALSE;
    inHoldPhase := FALSE;
    holdTimer(IN := FALSE, PT := T#500ms);
    THICKNESS_ALARM := FALSE;
END_IF;

(* When VALID is FALSE, ensure alarm and timer are cleared *)
IF NOT THICKNESS_SIGNAL_VALID THEN
    latch := FALSE;
    inHoldPhase := FALSE;
    holdTimer(IN := FALSE, PT := T#500ms);
    THICKNESS_ALARM := FALSE;
END_IF;

(* Process fault: activate alarm and record history *)
IF faultRising.Q THEN
    Slab_Fault_Counter := Slab_Fault_Counter + 1;

    FOR tmpI := 4 TO 1 BY -1 DO
        Slab_Fault_History[tmpI] := Slab_Fault_History[tmpI - 1];
    END_FOR;

    Slab_Fault_History[0] := FaultTimestamp;

    latch := TRUE;
    inHoldPhase := TRUE;
    holdTimer(IN := FALSE, PT := T#500ms);
    holdTimer(IN := TRUE, PT := T#500ms);
    THICKNESS_ALARM := TRUE;
END_IF;

(* Alarm follows latch during hold phase, then follows fault *)
IF latch THEN
    IF inHoldPhase THEN
        THICKNESS_ALARM := TRUE;
    ELSE
        THICKNESS_ALARM := THICKNESS_FAULT;
    END_IF;
ELSE
    THICKNESS_ALARM := FALSE;
END_IF;

(* Update hold phase and timer *)
IF inHoldPhase THEN
    IF holdTimer.Q THEN
        inHoldPhase := FALSE;
        IF NOT THICKNESS_FAULT THEN
            latch := FALSE;
        END_IF;
    END_IF;
END_IF;

(* Accumulate runtime while cutting normally *)
IF CUTTING_RUN AND THICKNESS_SIGNAL_VALID AND NOT THICKNESS_FAULT THEN
    Slab_Runtime_Accumulator := Slab_Runtime_Accumulator + TO_LTIME(CycleTime);
END_IF;

(* Update previous state for edge detection *)
prevFault := THICKNESS_FAULT;
prevValid := THICKNESS_SIGNAL_VALID;

END_FUNCTION_BLOCK

(* ---- public-medium-06.candidate_04.st ---- *)
FUNCTION_BLOCK SlabThicknessMonitor
VAR_INPUT
    THICKNESS_FAULT        : BOOL;
    THICKNESS_SIGNAL_VALID : BOOL;
    CUTTING_RUN            : BOOL;
    FaultTimestamp         : DINT;
    CycleTime              : TIME;
END_VAR

VAR_OUTPUT
    THICKNESS_ALARM          : BOOL;
    Slab_Fault_Counter       : UINT;
    Slab_Runtime_Accumulator : LTIME;
    Slab_Fault_History       : ARRAY[0..4] OF DINT;
END_VAR

VAR
    faultRising  : R_TRIG;
    validFalling : R_TRIG;
    prevFault    : BOOL;
    prevValid    : BOOL;
    holdTimer    : TON;
    holdActive   : BOOL;
    tmpI         : UINT;
END_VAR

(* ENGINEERING_CONTRACT
 * ┌─────────────────────────────────────────────────────────────────────────────────────────────┐
 * │ OUTPUT STATE TABLE                                                                           │
 * ├─────────────────┬───────────────────────────────────────────────────────────────────────────┤
 * │ THICKNESS_ALARM │ Activation:   immediate on FALSE-to-TRUE of FAULT while VALID=TRUE        │
 * │                 │ Retention:    holds TRUE for >= 500ms; then follows FAULT (PUB001)       │
 * │                 │ Reset:        VALID=FALSE clears alarm+hold; power-up clears (PUB004)    │
 * │                 │ Same-scan:    on VALID=FALSE, alarm OFF immediately; holdActive cleared  │
 * ├─────────────────┼───────────────────────────────────────────────────────────────────────────┤
 * │ Slab_Fault_     │ Activation:   FALSE-to-TRUE of FAULT while VALID=TRUE (PUB002)            │
 * │ Counter         │ Retention:    monotonically increasing; never auto-decremented           │
 * │                 │ Reset:        power-up only (PUB005)                                     │
 * ├─────────────────┼───────────────────────────────────────────────────────────────────────────┤
 * │ Slab_Runtime_   │ Activation:   CUTTING_RUN AND VALID AND NOT FAULT each scan (PUB003)     │
 * │ Accumulator     │ Retention:    preserved when conditions not met                          │
 * │                 │ Reset:        power-up only (PUB005)                                     │
 * │                 │ Units:        LTIME nanoseconds; CycleTime TIME converted via TO_LTIME   │
 * ├─────────────────┼───────────────────────────────────────────────────────────────────────────┤
 * │ Slab_Fault_     │ Activation:   new entry at index 0 on valid fault transition (PUB002)    │
 * │ History[0..4]   │ Shift:        older entries shift toward higher indices (PUB002)          │
 * │                 │ Retention:    five most recent; read-only to callers (PUB005)            │
 * │                 │ Reset:        power-up only (PUB005)                                     │
 * └─────────────────┴───────────────────────────────────────────────────────────────────────────┘
 *
 * ┌─────────────────────────────────────────────────────────────────────────────────────────────┐
 * │ TIMING BOUNDARY (PUB001)                                                                    │
 * │ - 500ms minimum hold: TON.Q = elapsed >= PT; first satisfying tick = 500 ticks @ 1ms       │
 * │ - holdActive ensures timer runs exactly once per fault; no continuous re-triggering        │
 * └─────────────────────────────────────────────────────────────────────────────────────────────┘
 *
 * CONTRACT_RULES []
 *)

(* Power-up initialization: VAR initial values handle all state to zero *)

(* Detect rising edge of fault while signal is valid *)
faultRising(CLK := THICKNESS_SIGNAL_VALID AND THICKNESS_FAULT AND NOT prevFault);

(* Detect falling edge of VALID *)
validFalling(CLK := prevValid AND NOT THICKNESS_SIGNAL_VALID);

(* Clear alarm and hold state when signal lost or invalidated *)
IF validFalling.Q OR NOT THICKNESS_SIGNAL_VALID THEN
    THICKNESS_ALARM := FALSE;
    holdActive      := FALSE;
    holdTimer(IN := FALSE, PT := T#500ms);
END_IF;

(* Process new fault: activate alarm and start 500ms hold timer *)
IF faultRising.Q THEN
    Slab_Fault_Counter := Slab_Fault_Counter + 1;

    FOR tmpI := 4 TO 1 BY -1 DO
        Slab_Fault_History[tmpI] := Slab_Fault_History[tmpI - 1];
    END_FOR;
    Slab_Fault_History[0] := FaultTimestamp;

    THICKNESS_ALARM := TRUE;
    holdActive      := TRUE;
    holdTimer(IN := TRUE, PT := T#500ms);
END_IF;

(* After 500ms hold completes, let alarm follow fault state *)
IF holdTimer.Q AND holdActive THEN
    holdActive := FALSE;
    holdTimer(IN := FALSE, PT := T#500ms);
    THICKNESS_ALARM := THICKNESS_FAULT AND THICKNESS_SIGNAL_VALID;
END_IF;

(* Accumulate normal-cutting runtime *)
IF CUTTING_RUN AND THICKNESS_SIGNAL_VALID AND NOT THICKNESS_FAULT THEN
    Slab_Runtime_Accumulator := Slab_Runtime_Accumulator + TO_LTIME(CycleTime);
END_IF;

(* Update previous state for next-scan edge detection *)
prevFault := THICKNESS_FAULT;
prevValid := THICKNESS_SIGNAL_VALID;

END_FUNCTION_BLOCK

(* ---- public-medium-06.raw_candidate_01.st ---- *)
FUNCTION_BLOCK SlabThicknessMonitor
VAR_INPUT
    THICKNESS_FAULT        : BOOL;
    THICKNESS_SIGNAL_VALID : BOOL;
    CUTTING_RUN            : BOOL;
    FaultTimestamp         : DINT;
    CycleTime              : TIME;
END_VAR

VAR_OUTPUT
    THICKNESS_ALARM          : BOOL;
    Slab_Fault_Counter       : UINT;
    Slab_Runtime_Accumulator : LTIME;
    Slab_Fault_History       : ARRAY[0..4] OF DINT;
END_VAR

VAR
    faultRising      : R_TRIG;
    validFalling     : R_TRIG;
    prevFault        : BOOL;
    prevValid        : BOOL;
    holdTimer        : TON;
    tmpI             : UINT;
END_VAR

(* ENGINEERING_CONTRACT
 * ┌─────────────────────────────────────────────────────────────────────────────────────────────┐
 * │ OUTPUT STATE TABLE                                                                           │
 * ├─────────────────┬───────────────────────────────────────────────────────────────────────────┤
 * │ THICKNESS_ALARM │ Activation:   rising edge of THICKNESS_FAULT while VALID=TRUE (PUB001)    │
 * │                 │ Retention:    held >= 500 ms via TON; remains TRUE while FAULT persists   │
 * │                 │ Reset:        VALID=FALSE or power-up clears alarm and holding state (PUB004)│
 * │                 │ Same-scan:    if VALID drops mid-scan, alarm OFF regardless of FAULT state│
 * ├─────────────────┼───────────────────────────────────────────────────────────────────────────┤
 * │ Slab_Fault_     │ Activation:   FALSE-to-TRUE of FAULT while VALID=TRUE (PUB002)             │
 * │ Counter         │ Retention:    monotonically increasing; never auto-decremented             │
 * │                 │ Reset:        power-up only (PUB005); external callers cannot modify       │
 * │                 │ Boundary:     UINT range; overflow wraps per IEC 61131-3                  │
 * ├─────────────────┼───────────────────────────────────────────────────────────────────────────┤
 * │ Slab_Runtime_   │ Activation:   CUTTING_RUN AND VALID AND NOT FAULT each scan (PUB003)       │
 * │ Accumulator     │ Retention:    preserved when conditions not met; never auto-cleared       │
 * │                 │ Reset:        power-up only (PUB005); uses LTIME nanoseconds internally   │
 * │                 │ Units:        CycleTime (TIME/ms) converted to LTIME (ns) before add      │
 * ├─────────────────┼───────────────────────────────────────────────────────────────────────────┤
 * │ Slab_Fault_     │ Activation:   new entry at index 0 on valid fault transition (PUB002)     │
 * │ History[0..4]   │ Shift:        older entries shift toward higher indices (PUB002)           │
 * │                 │ Retention:    five most recent; older beyond index 4 are discarded        │
 * │                 │ Reset:        power-up zeros all five entries (PUB005); read-only to callers│
 * └─────────────────┴───────────────────────────────────────────────────────────────────────────┘
 *
 * ┌─────────────────────────────────────────────────────────────────────────────────────────────┐
 * │ INPUT BEHAVIOR                                                                               │
 * ├───────────────────────────────┬─────────────────────────────────────────────────────────────┤
 * │ THICKNESS_SIGNAL_VALID=FALSE  │ alarm OFF, timer reset, no fault record, no runtime accum   │
 * │ THICKNESS_SIGNAL_VALID=TRUE   │ normal monitoring; alarm follows FAULT, counter/hist update │
 * │ CUTTING_RUN=FALSE             │ no runtime accumulation (fault monitoring still active)     │
 * │ CycleTime positive assumption │ caller guarantees > T#0s per task spec                     │
 * └───────────────────────────────┴─────────────────────────────────────────────────────────────┘
 *
 * ┌─────────────────────────────────────────────────────────────────────────────────────────────┐
 * │ TIMING BOUNDARY (PUB001, PUB003)                                                            │
 * │ - 500 ms hold: TON.Q = elapsed >= PT; first satisfying tick = ceil(500ms/1ms) = 500 ticks   │
 * │ - No implicit one-scan delay; timer enable and Q check occur in same invocation            │
 * └─────────────────────────────────────────────────────────────────────────────────────────────┘
 *
 * CONTRACT_RULES [{"kind": "hold_until_reset", "output": "THICKNESS_ALARM", "set_input": "THICKNESS_FAULT", "reset_input": null}]
 *)

(* Power-up initialization: handled by VAR initial values *)

(* Detect rising edge of fault while signal is valid *)
faultRising(CLK := THICKNESS_FAULT AND THICKNESS_SIGNAL_VALID AND NOT prevFault);

(* Detect falling edge of VALID to clear alarm and timer *)
validFalling(CLK := prevValid AND NOT THICKNESS_SIGNAL_VALID);

(* Handle signal invalidation: clear alarm and timer holding state *)
IF validFalling.Q THEN
    THICKNESS_ALARM := FALSE;
    holdTimer(IN := FALSE, PT := T#500ms);
END_IF

(* When VALID is FALSE, ensure alarm and timer are cleared *)
IF NOT THICKNESS_SIGNAL_VALID THEN
    THICKNESS_ALARM := FALSE;
    holdTimer(IN := FALSE, PT := T#500ms);
END_IF

(* Process fault: activate alarm and record history *)
IF faultRising.Q THEN
    (* Increment fault counter *)
    Slab_Fault_Counter := Slab_Fault_Counter + 1;

    (* Shift history: move entries toward higher indices *)
    FOR tmpI := 4 TO 1 BY -1 DO
        Slab_Fault_History[tmpI] := Slab_Fault_History[tmpI - 1];
    END_FOR;

    (* Store new fault timestamp at index 0 *)
    Slab_Fault_History[0] := FaultTimestamp;

    (* Activate alarm and start hold timer *)
    THICKNESS_ALARM := TRUE;
    holdTimer(IN := TRUE, PT := T#500ms);
END_IF;

(* Maintain alarm while fault persists (after initial 500ms hold) *)
IF holdTimer.Q THEN
    THICKNESS_ALARM := THICKNESS_FAULT AND THICKNESS_SIGNAL_VALID;
    holdTimer(IN := THICKNESS_ALARM, PT := T#500ms);
END_IF;

(* Accumulate runtime while cutting normally *)
IF CUTTING_RUN AND THICKNESS_SIGNAL_VALID AND NOT THICKNESS_FAULT THEN
    Slab_Runtime_Accumulator := Slab_Runtime_Accumulator + TO_LTIME(CycleTime);
END_IF;

(* Update previous state for edge detection on next scan *)
prevFault := THICKNESS_FAULT;
prevValid := THICKNESS_SIGNAL_VALID;

END_FUNCTION_BLOCK

(* ---- public-medium-06.raw_candidate_02.st ---- *)
FUNCTION_BLOCK SlabThicknessMonitor
VAR_INPUT
    THICKNESS_FAULT        : BOOL;
    THICKNESS_SIGNAL_VALID : BOOL;
    CUTTING_RUN            : BOOL;
    FaultTimestamp         : DINT;
    CycleTime              : TIME;
END_VAR

VAR_OUTPUT
    THICKNESS_ALARM          : BOOL;
    Slab_Fault_Counter       : UINT;
    Slab_Runtime_Accumulator : LTIME;
    Slab_Fault_History       : ARRAY[0..4] OF DINT;
END_VAR

VAR
    faultRising : R_TRIG;
    prevFault   : BOOL;
    prevValid   : BOOL;
    holdTimer   : TON;
    tmpI        : UINT;
END_VAR

(* ENGINEERING_CONTRACT
 * ┌─────────────────────────────────────────────────────────────────────────────────────────────┐
 * │ OUTPUT STATE TABLE                                                                           │
 * ├─────────────────┬───────────────────────────────────────────────────────────────────────────┤
 * │ THICKNESS_ALARM │ Activation:   immediate on rising edge of FAULT while VALID=TRUE (PUB001) │
 * │                 │ Retention:    hold >= 500ms via TON after FAULT drops; persists if FAULT │
 * │                 │               remains TRUE                                                │
 * │                 │ Reset:        VALID=FALSE clears alarm and timer holding state (PUB004)   │
 * │                 │ Same-scan:    alarm OFF immediately when VALID drops                      │
 * ├─────────────────┼───────────────────────────────────────────────────────────────────────────┤
 * │ Slab_Fault_     │ Activation:   FALSE-to-TRUE of FAULT while VALID=TRUE (PUB002)            │
 * │ Counter         │ Retention:    monotonically increasing; never auto-decremented            │
 * │                 │ Reset:        power-up only (PUB005)                                      │
 * │                 │ Boundary:     UINT range                                                  │
 * ├─────────────────┼───────────────────────────────────────────────────────────────────────────┤
 * │ Slab_Runtime_   │ Activation:   CUTTING_RUN AND VALID AND NOT FAULT AND NOT faultRising     │
 * │ Accumulator     │               (excludes scan where fault just transitioned TRUE) (PUB003) │
 * │                 │ Retention:    preserved when conditions not met                           │
 * │                 │ Reset:        power-up only (PUB005)                                      │
 * │                 │ Units:        CycleTime converted to LTIME ns before add                  │
 * ├─────────────────┼───────────────────────────────────────────────────────────────────────────┤
 * │ Slab_Fault_     │ Activation:   new entry at index 0 on valid fault transition (PUB002)     │
 * │ History[0..4]   │ Shift:        older entries shift toward higher indices (PUB002)          │
 * │                 │ Retention:    five most recent; older beyond index 4 discarded            │
 * │                 │ Reset:        power-up zeros all five entries (PUB005)                    │
 * └─────────────────┴───────────────────────────────────────────────────────────────────────────┘
 *
 * ┌─────────────────────────────────────────────────────────────────────────────────────────────┐
 * │ TIMING BOUNDARY (PUB001)                                                                    │
 * │ - 500ms hold: TON.Q = elapsed >= PT; first satisfying tick = 500 ticks at 1ms quantum      │
 * │ - Alarm reactivates immediately via R_TRIG on same-scan FAULT transitions                  │
 * │ - Timer resets when alarm deactivates to prevent stale elapsed time                        │
 * └─────────────────────────────────────────────────────────────────────────────────────────────┘
 *
 * CONTRACT_RULES [{"kind": "hold_until_reset", "output": "THICKNESS_ALARM", "set_input": "THICKNESS_FAULT", "reset_input": null}]
 *)

(* Power-up initialization: VAR initial values handle zeroing *)

(* Detect rising edge of fault while signal is valid *)
faultRising(CLK := THICKNESS_FAULT AND THICKNESS_SIGNAL_VALID AND NOT prevFault);

(* Clear alarm and timer when signal becomes invalid *)
IF NOT THICKNESS_SIGNAL_VALID THEN
    THICKNESS_ALARM := FALSE;
    holdTimer(IN := FALSE, PT := T#500ms);
END_IF;

(* Activate alarm immediately on valid fault rising edge *)
IF faultRising.Q THEN
    THICKNESS_ALARM := TRUE;
    holdTimer(IN := TRUE, PT := T#500ms);
END_IF;

(* Maintain alarm while fault persists after initial hold *)
IF holdTimer.Q THEN
    THICKNESS_ALARM := THICKNESS_FAULT AND THICKNESS_SIGNAL_VALID;
    holdTimer(IN := THICKNESS_ALARM, PT := T#500ms);
END_IF;

(* Record fault: increment counter and shift history *)
IF faultRising.Q THEN
    Slab_Fault_Counter := Slab_Fault_Counter + 1;
    FOR tmpI := 4 TO 1 BY -1 DO
        Slab_Fault_History[tmpI] := Slab_Fault_History[tmpI - 1];
    END_FOR;
    Slab_Fault_History[0] := FaultTimestamp;
END_IF;

(* Accumulate runtime only while cutting normally (excludes fault-transition scan) *)
IF CUTTING_RUN AND THICKNESS_SIGNAL_VALID AND NOT THICKNESS_FAULT AND NOT faultRising.Q THEN
    Slab_Runtime_Accumulator := Slab_Runtime_Accumulator + TO_LTIME(CycleTime);
END_IF;

(* Update previous state for edge detection *)
prevFault := THICKNESS_FAULT;
prevValid := THICKNESS_SIGNAL_VALID;

END_FUNCTION_BLOCK

(* ---- public-medium-06.raw_candidate_03.st ---- *)
FUNCTION_BLOCK SlabThicknessMonitor
VAR_INPUT
    THICKNESS_FAULT        : BOOL;
    THICKNESS_SIGNAL_VALID : BOOL;
    CUTTING_RUN            : BOOL;
    FaultTimestamp         : DINT;
    CycleTime              : TIME;
END_VAR

VAR_OUTPUT
    THICKNESS_ALARM          : BOOL;
    Slab_Fault_Counter       : UINT;
    Slab_Runtime_Accumulator : LTIME;
    Slab_Fault_History       : ARRAY[0..4] OF DINT;
END_VAR

VAR
    faultRising  : R_TRIG;
    validFalling : F_TRIG;
    prevFault    : BOOL;
    prevValid    : BOOL;
    holdTimer    : TON;
    latch        : BOOL;
    inHoldPhase  : BOOL;
    tmpI         : UINT;
END_VAR

(* ENGINEERING_CONTRACT
 * ┌─────────────────────────────────────────────────────────────────────────────────────────────┐
 * │ OUTPUT STATE TABLE                                                                           │
 * ├─────────────────┬───────────────────────────────────────────────────────────────────────────┤
 * │ THICKNESS_ALARM │ Activation:   immediate on rising edge of FAULT while VALID=TRUE (PUB001) │
 * │                 │ Retention:    held >= 500ms via TON; remains TRUE while FAULT persists   │
 * │                 │ Reset:        VALID=FALSE clears latch and timer (PUB004)                 │
 * │                 │ Same-scan:    latch set and timer started in same invocation as rising edge│
 * ├─────────────────┼───────────────────────────────────────────────────────────────────────────┤
 * │ Slab_Fault_     │ Activation:   FALSE-to-TRUE of FAULT while VALID=TRUE (PUB002)            │
 * │ Counter         │ Retention:    monotonically increasing; never auto-decremented            │
 * │                 │ Reset:        power-up only (PUB005)                                     │
 * │                 │ Boundary:     UINT range; overflow wraps per IEC 61131-3                 │
 * ├─────────────────┼───────────────────────────────────────────────────────────────────────────┤
 * │ Slab_Runtime_   │ Activation:   CUTTING_RUN AND VALID AND NOT FAULT each scan (PUB003)      │
 * │ Accumulator     │ Retention:    preserved when conditions not met; never auto-cleared      │
 * │                 │ Reset:        power-up only (PUB005)                                     │
 * │                 │ Units:        CycleTime (TIME) converted to LTIME (ns) before add        │
 * ├─────────────────┼───────────────────────────────────────────────────────────────────────────┤
 * │ Slab_Fault_     │ Activation:   new entry at index 0 on valid fault transition (PUB002)    │
 * │ History[0..4]   │ Shift:        older entries shift toward higher indices (PUB002)          │
 * │                 │ Retention:    five most recent; older beyond index 4 are discarded       │
 * │                 │ Reset:        power-up zeros all five entries (PUB005)                   │
 * └─────────────────┴───────────────────────────────────────────────────────────────────────────┘
 *
 * ┌─────────────────────────────────────────────────────────────────────────────────────────────┐
 * │ TIMING BOUNDARY (PUB001)                                                                    │
 * │ - 500 ms hold: TON.Q = elapsed >= PT; first satisfying tick = ceil(500ms/1ms) = 500 ticks  │
 * │ - Timer reset before restart ensures deterministic restart behavior                        │
 * └─────────────────────────────────────────────────────────────────────────────────────────────┘
 *
 * CONTRACT_RULES [{"kind": "hold_until_reset", "output": "THICKNESS_ALARM", "set_input": "THICKNESS_FAULT", "reset_input": null}]
 *)

(* Detect rising edge of fault while signal is valid *)
faultRising(CLK := THICKNESS_FAULT AND THICKNESS_SIGNAL_VALID AND NOT prevFault);

(* Detect falling edge of VALID to clear state *)
validFalling(CLK := prevValid AND NOT THICKNESS_SIGNAL_VALID);

(* Handle signal invalidation: clear latch, alarm, and timer *)
IF validFalling.Q THEN
    latch := FALSE;
    inHoldPhase := FALSE;
    holdTimer(IN := FALSE, PT := T#500ms);
    THICKNESS_ALARM := FALSE;
END_IF;

(* When VALID is FALSE, ensure alarm and timer are cleared *)
IF NOT THICKNESS_SIGNAL_VALID THEN
    latch := FALSE;
    inHoldPhase := FALSE;
    holdTimer(IN := FALSE, PT := T#500ms);
    THICKNESS_ALARM := FALSE;
END_IF;

(* Process fault: activate alarm and record history *)
IF faultRising.Q THEN
    Slab_Fault_Counter := Slab_Fault_Counter + 1;

    FOR tmpI := 4 TO 1 BY -1 DO
        Slab_Fault_History[tmpI] := Slab_Fault_History[tmpI - 1];
    END_FOR;

    Slab_Fault_History[0] := FaultTimestamp;

    latch := TRUE;
    inHoldPhase := TRUE;
    holdTimer(IN := FALSE, PT := T#500ms);
    holdTimer(IN := TRUE, PT := T#500ms);
    THICKNESS_ALARM := TRUE;
END_IF;

(* Alarm follows latch during hold phase, then follows fault *)
IF latch THEN
    IF inHoldPhase THEN
        THICKNESS_ALARM := TRUE;
    ELSE
        THICKNESS_ALARM := THICKNESS_FAULT;
    END_IF;
ELSE
    THICKNESS_ALARM := FALSE;
END_IF;

(* Update hold phase and timer *)
IF inHoldPhase THEN
    IF holdTimer.Q THEN
        inHoldPhase := FALSE;
        IF NOT THICKNESS_FAULT THEN
            latch := FALSE;
        END_IF;
    END_IF;
END_IF;

(* Accumulate runtime while cutting normally *)
IF CUTTING_RUN AND THICKNESS_SIGNAL_VALID AND NOT THICKNESS_FAULT THEN
    Slab_Runtime_Accumulator := Slab_Runtime_Accumulator + TO_LTIME(CycleTime);
END_IF;

(* Update previous state for edge detection *)
prevFault := THICKNESS_FAULT;
prevValid := THICKNESS_SIGNAL_VALID;

END_FUNCTION_BLOCK

(* ---- public-medium-06.raw_candidate_04.st ---- *)
FUNCTION_BLOCK SlabThicknessMonitor
VAR_INPUT
    THICKNESS_FAULT        : BOOL;
    THICKNESS_SIGNAL_VALID : BOOL;
    CUTTING_RUN            : BOOL;
    FaultTimestamp         : DINT;
    CycleTime              : TIME;
END_VAR

VAR_OUTPUT
    THICKNESS_ALARM          : BOOL;
    Slab_Fault_Counter       : UINT;
    Slab_Runtime_Accumulator : LTIME;
    Slab_Fault_History       : ARRAY[0..4] OF DINT;
END_VAR

VAR
    faultRising  : R_TRIG;
    validFalling : R_TRIG;
    prevFault    : BOOL;
    prevValid    : BOOL;
    holdTimer    : TON;
    holdActive   : BOOL;
    tmpI         : UINT;
END_VAR

(* ENGINEERING_CONTRACT
 * ┌─────────────────────────────────────────────────────────────────────────────────────────────┐
 * │ OUTPUT STATE TABLE                                                                           │
 * ├─────────────────┬───────────────────────────────────────────────────────────────────────────┤
 * │ THICKNESS_ALARM │ Activation:   immediate on FALSE-to-TRUE of FAULT while VALID=TRUE        │
 * │                 │ Retention:    holds TRUE for >= 500ms; then follows FAULT (PUB001)       │
 * │                 │ Reset:        VALID=FALSE clears alarm+hold; power-up clears (PUB004)    │
 * │                 │ Same-scan:    on VALID=FALSE, alarm OFF immediately; holdActive cleared  │
 * ├─────────────────┼───────────────────────────────────────────────────────────────────────────┤
 * │ Slab_Fault_     │ Activation:   FALSE-to-TRUE of FAULT while VALID=TRUE (PUB002)            │
 * │ Counter         │ Retention:    monotonically increasing; never auto-decremented           │
 * │                 │ Reset:        power-up only (PUB005)                                     │
 * ├─────────────────┼───────────────────────────────────────────────────────────────────────────┤
 * │ Slab_Runtime_   │ Activation:   CUTTING_RUN AND VALID AND NOT FAULT each scan (PUB003)     │
 * │ Accumulator     │ Retention:    preserved when conditions not met                          │
 * │                 │ Reset:        power-up only (PUB005)                                     │
 * │                 │ Units:        LTIME nanoseconds; CycleTime TIME converted via TO_LTIME   │
 * ├─────────────────┼───────────────────────────────────────────────────────────────────────────┤
 * │ Slab_Fault_     │ Activation:   new entry at index 0 on valid fault transition (PUB002)    │
 * │ History[0..4]   │ Shift:        older entries shift toward higher indices (PUB002)          │
 * │                 │ Retention:    five most recent; read-only to callers (PUB005)            │
 * │                 │ Reset:        power-up only (PUB005)                                     │
 * └─────────────────┴───────────────────────────────────────────────────────────────────────────┘
 *
 * ┌─────────────────────────────────────────────────────────────────────────────────────────────┐
 * │ TIMING BOUNDARY (PUB001)                                                                    │
 * │ - 500ms minimum hold: TON.Q = elapsed >= PT; first satisfying tick = 500 ticks @ 1ms       │
 * │ - holdActive ensures timer runs exactly once per fault; no continuous re-triggering        │
 * └─────────────────────────────────────────────────────────────────────────────────────────────┘
 *
 * CONTRACT_RULES []
 *)

(* Power-up initialization: VAR initial values handle all state to zero *)

(* Detect rising edge of fault while signal is valid *)
faultRising(CLK := THICKNESS_SIGNAL_VALID AND THICKNESS_FAULT AND NOT prevFault);

(* Detect falling edge of VALID *)
validFalling(CLK := prevValid AND NOT THICKNESS_SIGNAL_VALID);

(* Clear alarm and hold state when signal lost or invalidated *)
IF validFalling.Q OR NOT THICKNESS_SIGNAL_VALID THEN
    THICKNESS_ALARM := FALSE;
    holdActive      := FALSE;
    holdTimer(IN := FALSE, PT := T#500ms);
END_IF;

(* Process new fault: activate alarm and start 500ms hold timer *)
IF faultRising.Q THEN
    Slab_Fault_Counter := Slab_Fault_Counter + 1;

    FOR tmpI := 4 TO 1 BY -1 DO
        Slab_Fault_History[tmpI] := Slab_Fault_History[tmpI - 1];
    END_FOR;
    Slab_Fault_History[0] := FaultTimestamp;

    THICKNESS_ALARM := TRUE;
    holdActive      := TRUE;
    holdTimer(IN := TRUE, PT := T#500ms);
END_IF;

(* After 500ms hold completes, let alarm follow fault state *)
IF holdTimer.Q AND holdActive THEN
    holdActive := FALSE;
    holdTimer(IN := FALSE, PT := T#500ms);
    THICKNESS_ALARM := THICKNESS_FAULT AND THICKNESS_SIGNAL_VALID;
END_IF;

(* Accumulate normal-cutting runtime *)
IF CUTTING_RUN AND THICKNESS_SIGNAL_VALID AND NOT THICKNESS_FAULT THEN
    Slab_Runtime_Accumulator := Slab_Runtime_Accumulator + TO_LTIME(CycleTime);
END_IF;

(* Update previous state for next-scan edge detection *)
prevFault := THICKNESS_FAULT;
prevValid := THICKNESS_SIGNAL_VALID;

END_FUNCTION_BLOCK

(* ---- public-medium-07.candidate_01.st ---- *)
(* ENGINEERING_CONTRACT
 * HVAC Multi-mode Energy-Saving Control - Design Table
 *
 * Output: SUPPLY_FAN_RUN (BOOL)
 *   - Activation:    30s TON delay when OCCUPANCY_DETECTED=TRUE AND HVAC_MODE_SELECTOR<>3
 *   - Retention:     Holds TRUE once elapsed >= 30s until deactivated
 *   - Reset:         Immediate deactivation when OCCUPANCY_DETECTED=FALSE OR HVAC_MODE_SELECTOR=3
 *   - Same-scan:     Evaluate conditions before TON, update outputs after TON
 *   - Units:         30 seconds, TON.ET saturates at PT
 *
 * Output: TEMP_SETPOINT_ADJUST (INT, clamped ±4°C)
 *   - PUB001 §3: Auto mode - occupied: 0°C; unoccupied + energy_saving: +3°C; unoccupied + standard: +2°C
 *   - PUB002 §4: Comfort mode - occupied: 0°C; unoccupied: +1°C
 *   - PUB003 §5: Economy mode - occupied: 0°C; unoccupied: +4°C
 *   - PUB004 §6: Night mode (3) - +4°C regardless of occupancy
 *   - Retention:   Updated every scan from current inputs; no state retention between scans
 *   - Boundaries:  Clamped to [-4, +4] inclusive
 *
 * Initialization:
 *   - SUPPLY_FAN_RUN := FALSE on power-up (PUB006)
 *   - TEMP_SETPOINT_ADJUST := 0 on power-up (PUB006)
 *   - Timer state initialized by TON at first call (implicit)
 *
 * Edge Cases:
 *   - Night mode selected: fan disabled immediately, no delay (PUB001)
 *   - Occupancy lost: fan disabled immediately, timer reset (PUB001)
 *   - Recovery: full 30s delay required again (PUB001)
 *   - HVAC_MODE_SELECTOR values 0-3 only; caller supplies valid value
 *)

(* CONTRACT_RULES [] *)

FUNCTION_BLOCK HVAC_MultiMode_Control
VAR_INPUT
    OCCUPANCY_DETECTED  : BOOL;
    ENERGY_SAVING_MODE  : BOOL;
    HVAC_MODE_SELECTOR  : INT;
END_VAR

VAR_OUTPUT
    SUPPLY_FAN_RUN      : BOOL := FALSE;
    TEMP_SETPOINT_ADJUST : INT := 0;
END_VAR

VAR
    FanDelayTimer : TON;
    prevOccupancy : BOOL := FALSE;
    tmpOccupied   : BOOL;
    tmpFanEnable  : BOOL;
    tmpAdjust     : INT;
END_VAR

(* Same-scan logic: determine conditions before timer, then act *)
tmpOccupied := OCCUPANCY_DETECTED AND (HVAC_MODE_SELECTOR <> 3);

(* Fan enable request: occupied AND not night mode *)
tmpFanEnable := tmpOccupied;

(* Manage fan delay timer *)
IF tmpFanEnable THEN
    FanDelayTimer(IN := TRUE, PT := T#30S);
    (* TON.Q is TRUE when elapsed >= PT; TON.ET saturates at PT *)
    SUPPLY_FAN_RUN := FanDelayTimer.Q;
ELSE
    FanDelayTimer(IN := FALSE, PT := T#30S);
    SUPPLY_FAN_RUN := FALSE;
END_IF;

(* Temperature setpoint adjustment per mode *)
CASE HVAC_MODE_SELECTOR OF
    0: (* Auto mode *)
        IF OCCUPANCY_DETECTED THEN
            tmpAdjust := 0;
        ELSE
            IF ENERGY_SAVING_MODE THEN
                tmpAdjust := 3;
            ELSE
                tmpAdjust := 2;
            END_IF;
        END_IF;

    1: (* Comfort mode *)
        IF OCCUPANCY_DETECTED THEN
            tmpAdjust := 0;
        ELSE
            tmpAdjust := 1;
        END_IF;

    2: (* Economy mode *)
        IF OCCUPANCY_DETECTED THEN
            tmpAdjust := 0;
        ELSE
            tmpAdjust := 4;
        END_IF;

    3: (* Night mode *)
        tmpAdjust := 4;

    ELSE
        (* Fallback for invalid values; maintain last safe state *)
        tmpAdjust := 0;
END_CASE;

(* Clamp to ±4°C per PUB007 *)
IF tmpAdjust > 4 THEN
    tmpAdjust := 4;
ELSIF tmpAdjust < -4 THEN
    tmpAdjust := -4;
END_IF;

TEMP_SETPOINT_ADJUST := tmpAdjust;

(* Track occupancy for next scan *)
prevOccupancy := OCCUPANCY_DETECTED;

END_FUNCTION_BLOCK

(* ---- public-medium-07.raw_candidate_01.st ---- *)
(* ENGINEERING_CONTRACT
 * HVAC Multi-mode Energy-Saving Control - Design Table
 *
 * Output: SUPPLY_FAN_RUN (BOOL)
 *   - Activation:    30s TON delay when OCCUPANCY_DETECTED=TRUE AND HVAC_MODE_SELECTOR<>3
 *   - Retention:     Holds TRUE once elapsed >= 30s until deactivated
 *   - Reset:         Immediate deactivation when OCCUPANCY_DETECTED=FALSE OR HVAC_MODE_SELECTOR=3
 *   - Same-scan:     Evaluate conditions before TON, update outputs after TON
 *   - Units:         30 seconds, TON.ET saturates at PT
 *
 * Output: TEMP_SETPOINT_ADJUST (INT, clamped ±4°C)
 *   - PUB001 §3: Auto mode - occupied: 0°C; unoccupied + energy_saving: +3°C; unoccupied + standard: +2°C
 *   - PUB002 §4: Comfort mode - occupied: 0°C; unoccupied: +1°C
 *   - PUB003 §5: Economy mode - occupied: 0°C; unoccupied: +4°C
 *   - PUB004 §6: Night mode (3) - +4°C regardless of occupancy
 *   - Retention:   Updated every scan from current inputs; no state retention between scans
 *   - Boundaries:  Clamped to [-4, +4] inclusive
 *
 * Initialization:
 *   - SUPPLY_FAN_RUN := FALSE on power-up (PUB006)
 *   - TEMP_SETPOINT_ADJUST := 0 on power-up (PUB006)
 *   - Timer state initialized by TON at first call (implicit)
 *
 * Edge Cases:
 *   - Night mode selected: fan disabled immediately, no delay (PUB001)
 *   - Occupancy lost: fan disabled immediately, timer reset (PUB001)
 *   - Recovery: full 30s delay required again (PUB001)
 *   - HVAC_MODE_SELECTOR values 0-3 only; caller supplies valid value
 *)

(* CONTRACT_RULES [] *)

FUNCTION_BLOCK HVAC_MultiMode_Control
VAR_INPUT
    OCCUPANCY_DETECTED  : BOOL;
    ENERGY_SAVING_MODE  : BOOL;
    HVAC_MODE_SELECTOR  : INT;
END_VAR

VAR_OUTPUT
    SUPPLY_FAN_RUN      : BOOL := FALSE;
    TEMP_SETPOINT_ADJUST : INT := 0;
END_VAR

VAR
    FanDelayTimer : TON;
    prevOccupancy : BOOL := FALSE;
    tmpOccupied   : BOOL;
    tmpFanEnable  : BOOL;
    tmpAdjust     : INT;
END_VAR

(* Same-scan logic: determine conditions before timer, then act *)
tmpOccupied := OCCUPANCY_DETECTED AND (HVAC_MODE_SELECTOR <> 3);

(* Fan enable request: occupied AND not night mode *)
tmpFanEnable := tmpOccupied;

(* Manage fan delay timer *)
IF tmpFanEnable THEN
    FanDelayTimer(IN := TRUE, PT := T#30S);
    (* TON.Q is TRUE when elapsed >= PT; TON.ET saturates at PT *)
    SUPPLY_FAN_RUN := FanDelayTimer.Q;
ELSE
    FanDelayTimer(IN := FALSE, PT := T#30S);
    SUPPLY_FAN_RUN := FALSE;
END_IF;

(* Temperature setpoint adjustment per mode *)
CASE HVAC_MODE_SELECTOR OF
    0: (* Auto mode *)
        IF OCCUPANCY_DETECTED THEN
            tmpAdjust := 0;
        ELSE
            IF ENERGY_SAVING_MODE THEN
                tmpAdjust := 3;
            ELSE
                tmpAdjust := 2;
            END_IF;
        END_IF;

    1: (* Comfort mode *)
        IF OCCUPANCY_DETECTED THEN
            tmpAdjust := 0;
        ELSE
            tmpAdjust := 1;
        END_IF;

    2: (* Economy mode *)
        IF OCCUPANCY_DETECTED THEN
            tmpAdjust := 0;
        ELSE
            tmpAdjust := 4;
        END_IF;

    3: (* Night mode *)
        tmpAdjust := 4;

    ELSE
        (* Fallback for invalid values; maintain last safe state *)
        tmpAdjust := 0;
END_CASE;

(* Clamp to ±4°C per PUB007 *)
IF tmpAdjust > 4 THEN
    tmpAdjust := 4;
ELSIF tmpAdjust < -4 THEN
    tmpAdjust := -4;
END_IF;

TEMP_SETPOINT_ADJUST := tmpAdjust;

(* Track occupancy for next scan *)
prevOccupancy := OCCUPANCY_DETECTED;

END_FUNCTION_BLOCK

(* ---- public-medium-08.candidate_01.st ---- *)
(* ENGINEERING_CONTRACT
   PUB001: Parse dotted-decimal IPv4, validate 4 numeric segments 0-255
   PUB002: Network byte order assembly (MSB=first segment)
   PUB003: Invalid input → ipValue=0 (malformed, nondigit, wrong count, OOR)
   PUB004: Valid 0.0.0.0 also produces 0 (by assembly)

   State retention: None (stateless function block)
   Reset behavior: None (no reset input specified)
   First scan: Same as subsequent (no edge memory)
*)

(* CONTRACT_RULES [] *)

FUNCTION_BLOCK IPv4_Parse
VAR_INPUT
    ipText : STRING(254);
END_VAR
VAR_OUTPUT
    ipValue : UDINT := 0;
END_VAR
VAR
    tmp_pos : UDINT;
    tmp_seg_idx : UDINT;
    tmp_char : BYTE;
    tmp_seg_val : UDINT;
    tmp_result : UDINT;
END_VAR

tmp_pos := 0;
tmp_seg_idx := 0;
tmp_result := 0;
tmp_seg_val := 0;

WHILE tmp_pos < LEN(ipText) DO
    tmp_char := ipText[tmp_pos];

    IF tmp_char >= 48 AND tmp_char <= 57 THEN
        tmp_seg_val := tmp_seg_val * 10 + TO_UDINT(tmp_char - 48);

        IF tmp_seg_val > 255 THEN
            ipValue := 0;
            RETURN;
        END_IF;

        tmp_pos := tmp_pos + 1;

    ELSE

        IF tmp_seg_idx >= 3 THEN
            ipValue := 0;
            RETURN;
        END_IF;

        CASE tmp_seg_idx OF
            0: tmp_result := SHL(tmp_seg_val, 24);
            1: tmp_result := tmp_result OR SHL(tmp_seg_val, 16);
            2: tmp_result := tmp_result OR SHL(tmp_seg_val, 8);
            3: tmp_result := tmp_result OR tmp_seg_val;
        END_CASE;

        tmp_seg_idx := tmp_seg_idx + 1;
        tmp_seg_val := 0;

        IF tmp_pos < LEN(ipText) THEN
            tmp_pos := tmp_pos + 1;
        END_IF;
    END_IF;
END_WHILE;

IF tmp_seg_idx <> 3 THEN
    ipValue := 0;
ELSE
    tmp_result := tmp_result OR tmp_seg_val;
    ipValue := tmp_result;
END_IF;

END_FUNCTION_BLOCK

(* ---- public-medium-08.candidate_02.st ---- *)
(* ENGINEERING_CONTRACT
   PUB001: Parse dotted-decimal IPv4, validate 4 numeric segments 0-255
   PUB002: Network byte order assembly (MSB=first segment)
   PUB003: Invalid input → ipValue=0 (malformed, nondigit, wrong count, OOR)
   PUB004: Valid 0.0.0.0 also produces 0 (by assembly)

   Empty segment: rejected unless it's segment 0 with value 0 (0.0.0.0 case)
   State retention: None (stateless function block)
   Reset behavior: None (no reset input specified)
*)

(* CONTRACT_RULES [] *)

FUNCTION_BLOCK IPv4_Parse
VAR_INPUT
    ipText : STRING(254);
END_VAR
VAR_OUTPUT
    ipValue : UDINT := 0;
END_VAR
VAR
    tmp_pos : UDINT;
    tmp_seg_idx : UDINT;
    tmp_char : BYTE;
    tmp_seg_val : UDINT;
    tmp_result : UDINT;
END_VAR

tmp_pos := 0;
tmp_seg_idx := 0;
tmp_result := 0;
tmp_seg_val := 0;

WHILE tmp_pos < LEN(ipText) DO
    tmp_char := ipText[tmp_pos];

    IF tmp_char >= 48 AND tmp_char <= 57 THEN
        tmp_seg_val := tmp_seg_val * 10 + TO_UDINT(tmp_char - 48);

        IF tmp_seg_val > 255 THEN
            ipValue := 0;
            RETURN;
        END_IF;

        tmp_pos := tmp_pos + 1;

    ELSE

        IF tmp_seg_idx >= 3 THEN
            ipValue := 0;
            RETURN;
        END_IF;

        IF tmp_seg_val = 0 AND tmp_seg_idx < 3 THEN
            ipValue := 0;
            RETURN;
        END_IF;

        CASE tmp_seg_idx OF
            0: tmp_result := SHL(tmp_seg_val, 24);
            1: tmp_result := tmp_result OR SHL(tmp_seg_val, 16);
            2: tmp_result := tmp_result OR SHL(tmp_seg_val, 8);
            3: tmp_result := tmp_result OR tmp_seg_val;
        END_CASE;

        tmp_seg_idx := tmp_seg_idx + 1;
        tmp_seg_val := 0;

        IF tmp_pos < LEN(ipText) THEN
            tmp_pos := tmp_pos + 1;
        END_IF;
    END_IF;
END_WHILE;

IF tmp_seg_idx <> 3 THEN
    ipValue := 0;
ELSE
    tmp_result := tmp_result OR tmp_seg_val;
    ipValue := tmp_result;
END_IF;

END_FUNCTION_BLOCK

(* ---- public-medium-08.candidate_04.st ---- *)
(* ENGINEERING_CONTRACT
   PUB001: Parse dotted-decimal IPv4, validate 4 numeric segments 0-255
   PUB002: Network byte order assembly (MSB=first segment)
   PUB003: Invalid input → ipValue=0 (malformed, nondigit, wrong count, OOR)
   PUB004: Valid 0.0.0.0 also produces 0 (by assembly)

   State retention: None (stateless function block)
   Reset behavior: None (no reset input specified)
   First scan: Same as subsequent (no edge memory)

   Bug fix: Reject empty segments (consecutive delimiters like "1..2.3")
   by tracking nonempty digit accumulation per segment
*)

(* CONTRACT_RULES [] *)

FUNCTION_BLOCK IPv4_Parse
VAR_INPUT
    ipText : STRING(254);
END_VAR
VAR_OUTPUT
    ipValue : UDINT := 0;
END_VAR
VAR
    tmp_pos : UDINT;
    tmp_seg_idx : UDINT;
    tmp_char : BYTE;
    tmp_seg_val : UDINT;
    tmp_result : UDINT;
    tmp_seg_nonempty : BOOL;
END_VAR

tmp_pos := 0;
tmp_seg_idx := 0;
tmp_result := 0;
tmp_seg_val := 0;
tmp_seg_nonempty := FALSE;

WHILE tmp_pos < LEN(ipText) DO
    tmp_char := ipText[tmp_pos];

    IF tmp_char >= 48 AND tmp_char <= 57 THEN
        tmp_seg_val := tmp_seg_val * 10 + TO_UDINT(tmp_char - 48);

        IF tmp_seg_val > 255 THEN
            ipValue := 0;
            RETURN;
        END_IF;

        tmp_seg_nonempty := TRUE;
        tmp_pos := tmp_pos + 1;

    ELSIF tmp_char = 46 THEN

        IF NOT tmp_seg_nonempty THEN
            ipValue := 0;
            RETURN;
        END_IF;

        IF tmp_seg_idx >= 3 THEN
            ipValue := 0;
            RETURN;
        END_IF;

        CASE tmp_seg_idx OF
            0: tmp_result := SHL(tmp_seg_val, 24);
            1: tmp_result := tmp_result OR SHL(tmp_seg_val, 16);
            2: tmp_result := tmp_result OR SHL(tmp_seg_val, 8);
        END_CASE;

        tmp_seg_idx := tmp_seg_idx + 1;
        tmp_seg_val := 0;
        tmp_seg_nonempty := FALSE;
        tmp_pos := tmp_pos + 1;
    ELSE

        ipValue := 0;
        RETURN;
    END_IF;
END_WHILE;

IF tmp_seg_idx <> 3 THEN
    ipValue := 0;
ELSE
    tmp_result := tmp_result OR tmp_seg_val;
    ipValue := tmp_result;
END_IF;

END_FUNCTION_BLOCK

(* ---- public-medium-08.raw_candidate_01.st ---- *)
(* ENGINEERING_CONTRACT
   PUB001: Parse dotted-decimal IPv4, validate 4 numeric segments 0-255
   PUB002: Network byte order assembly (MSB=first segment)
   PUB003: Invalid input → ipValue=0 (malformed, nondigit, wrong count, OOR)
   PUB004: Valid 0.0.0.0 also produces 0 (by assembly)

   State retention: None (stateless function block)
   Reset behavior: None (no reset input specified)
   First scan: Same as subsequent (no edge memory)
*)

(* CONTRACT_RULES [] *)

FUNCTION_BLOCK IPv4_Parse
VAR_INPUT
    ipText : STRING(254);
END_VAR
VAR_OUTPUT
    ipValue : UDINT := 0;
END_VAR
VAR
    tmp_pos : UDINT;
    tmp_seg_idx : UDINT;
    tmp_char : BYTE;
    tmp_seg_val : UDINT;
    tmp_result : UDINT;
END_VAR

tmp_pos := 0;
tmp_seg_idx := 0;
tmp_result := 0;
tmp_seg_val := 0;

WHILE tmp_pos < LEN(ipText) DO
    tmp_char := ipText[tmp_pos];

    IF tmp_char >= 48 AND tmp_char <= 57 THEN
        tmp_seg_val := tmp_seg_val * 10 + TO_UDINT(tmp_char - 48);

        IF tmp_seg_val > 255 THEN
            ipValue := 0;
            RETURN;
        END_IF;

        tmp_pos := tmp_pos + 1;

    ELSE

        IF tmp_seg_idx >= 3 THEN
            ipValue := 0;
            RETURN;
        END_IF;

        CASE tmp_seg_idx OF
            0: tmp_result := SHL(tmp_seg_val, 24);
            1: tmp_result := tmp_result OR SHL(tmp_seg_val, 16);
            2: tmp_result := tmp_result OR SHL(tmp_seg_val, 8);
            3: tmp_result := tmp_result OR tmp_seg_val;
        END_CASE

        tmp_seg_idx := tmp_seg_idx + 1;
        tmp_seg_val := 0;

        IF tmp_pos < LEN(ipText) THEN
            tmp_pos := tmp_pos + 1;
        END_IF;
    END_IF;
END_WHILE;

IF tmp_seg_idx <> 3 THEN
    ipValue := 0;
ELSE
    tmp_result := tmp_result OR tmp_seg_val;
    ipValue := tmp_result;
END_IF;

END_FUNCTION_BLOCK

(* ---- public-medium-08.raw_candidate_02.st ---- *)
(* ENGINEERING_CONTRACT
   PUB001: Parse dotted-decimal IPv4, validate 4 numeric segments 0-255
   PUB002: Network byte order assembly (MSB=first segment)
   PUB003: Invalid input → ipValue=0 (malformed, nondigit, wrong count, OOR)
   PUB004: Valid 0.0.0.0 also produces 0 (by assembly)

   Empty segment: rejected unless it's segment 0 with value 0 (0.0.0.0 case)
   State retention: None (stateless function block)
   Reset behavior: None (no reset input specified)
*)

(* CONTRACT_RULES [] *)

FUNCTION_BLOCK IPv4_Parse
VAR_INPUT
    ipText : STRING(254);
END_VAR
VAR_OUTPUT
    ipValue : UDINT := 0;
END_VAR
VAR
    tmp_pos : UDINT;
    tmp_seg_idx : UDINT;
    tmp_char : BYTE;
    tmp_seg_val : UDINT;
    tmp_result : UDINT;
END_VAR

tmp_pos := 0;
tmp_seg_idx := 0;
tmp_result := 0;
tmp_seg_val := 0;

WHILE tmp_pos < LEN(ipText) DO
    tmp_char := ipText[tmp_pos];

    IF tmp_char >= 48 AND tmp_char <= 57 THEN
        tmp_seg_val := tmp_seg_val * 10 + TO_UDINT(tmp_char - 48);

        IF tmp_seg_val > 255 THEN
            ipValue := 0;
            RETURN;
        END_IF;

        tmp_pos := tmp_pos + 1;

    ELSE

        IF tmp_seg_idx >= 3 THEN
            ipValue := 0;
            RETURN;
        END_IF;

        IF tmp_seg_val = 0 AND tmp_seg_idx < 3 THEN
            ipValue := 0;
            RETURN;
        END_IF;

        CASE tmp_seg_idx OF
            0: tmp_result := SHL(tmp_seg_val, 24);
            1: tmp_result := tmp_result OR SHL(tmp_seg_val, 16);
            2: tmp_result := tmp_result OR SHL(tmp_seg_val, 8);
            3: tmp_result := tmp_result OR tmp_seg_val;
        END_CASE;

        tmp_seg_idx := tmp_seg_idx + 1;
        tmp_seg_val := 0;

        IF tmp_pos < LEN(ipText) THEN
            tmp_pos := tmp_pos + 1;
        END_IF;
    END_IF;
END_WHILE;

IF tmp_seg_idx <> 3 THEN
    ipValue := 0;
ELSE
    tmp_result := tmp_result OR tmp_seg_val;
    ipValue := tmp_result;
END_IF;

END_FUNCTION_BLOCK
